(* IEC 61131-3 sources: daoli-st-library/DL_Motion (part 5) *)

(* ---- FB_DL_AgvPathTrackSeq.st ---- *)
// FB_DL_AgvPathTrackSeq v1.0.0
// 开源溯源：clean-room 自研（族 DL_Motion，ST 生态实测 0 命中，无外部代码引入）
(*
  功能: AGV 路径跟踪序列相位机：IDLE →(xStart∧xEnable) ALIGN →(双容差对齐) TRACK
        →(xObstacle) AVOID →(障碍解除∧保持 2 s) TRACK；TRACK →(xDockZone) DOCK
        →(对齐∧dist<0.05) IDLE 置 xDone。速度按 0.5 m/s² 斜坡逼近（增量 0.5·fCycleS，不阶跃），
        AVOID 与 FAULT 相强制零速零转。几何律全部委托外部 FC，本件不含三角函数。
  邻件: 对桩律 FC_DL_AgvChargeDockAlignCalc、限速 FC_DL_AgvSpeedLimitProfileCalc 为上游计算件。
  码表: 9311 入参非有限｜9312 组态非法(fSpeedLimit/fCycleS≤0)｜9313 相超时(ALIGN 5s/AVOID 保持/DOCK 15s)
        9314 相位落 ELSE 兜底｜9315 信息级序列完成（不置故障）。故障码锁存至 xReset 上升沿。
  边界: 无方法块/无属性块/无全局变量/无物理 IO 地址；三 TON 单相独占且无条件刷新。
*)
TYPE E_DL_AgvTrackState :
(
    IDLE  := 0,     // 空闲：等启动指令 [-] / Idle, waiting start
    ALIGN := 10,    // 对准：横向与角度对桩 [-] / Aligning to dock
    TRACK := 20,    // 跟踪：沿路径行驶 [-] / Tracking the path
    AVOID := 30,    // 避障：零速等待障碍解除 [-] / Avoiding obstacle
    DOCK  := 40,    // 入桩：末端贴近充电桩 [-] / Docking approach
    FAULT := 90     // 故障：锁存，仅复位沿可出 [-] / Fault latched
);
END_TYPE
FUNCTION_BLOCK FB_DL_AgvPathTrackSeq
VAR_INPUT
    xEnable     : BOOL := FALSE;        // 使能，FALSE 时全相冻结 [-] / Enable gate
    xStart      : BOOL := FALSE;        // 启动指令，上升沿有效 [-] / Start rising edge
    xReset      : BOOL := FALSE;        // 复位，上升沿清故障锁存 [-] / Reset rising edge
    xObstacle   : BOOL := FALSE;        // 障碍检测输入 [-] / Obstacle detected
    xDockZone   : BOOL := FALSE;        // 入桩区检测输入 [-] / Dock zone detected
    fOffsetY    : REAL := 0.0;          // 横向偏差 [m]，左正 / Lateral offset [m]
    fAngleErr   : REAL := 0.0;          // 角度偏差 [rad]，左正 / Angular error [rad]
    fDist       : REAL := 2.0;          // 到桩距离 [m] / Distance to dock [m]
    fSpeedLimit : REAL := 1.0;          // 允许限速 [m/s]，域 > 0 / Speed limit [m/s]
    fCycleS     : REAL := 0.01;         // 任务周期 [s]，域 > 0 / Task cycle time [s]
END_VAR
VAR_OUTPUT
    eState      : E_DL_AgvTrackState;   // 相位出口，段尾单点映射 [-] / Phase outlet
    xRun        : BOOL;                 // 运行中标志（非 IDLE 非 FAULT）[-] / Running flag
    fSpeedCmd   : REAL;                 // 前进速度指令 [m/s] / Speed command [m/s]
    fYawRateCmd : REAL;                 // 转向角速度指令 [rad/s] / Yaw rate command [rad/s]
    xDone       : BOOL;                 // 序列完成单拍脉冲 [-] / Done one-shot pulse
    xFault      : BOOL;                 // 故障锁存标志 [-] / Fault latch flag
    uErrorId    : UDINT;                // 事件码，0 = 无事件 / Event code
END_VAR
VAR
    tonAlign  : TON;                    // ALIGN 相超时 5 s，单相独占刷新 / Align timeout
    tonAvoid  : TON;                    // AVOID 障碍保持窗 2 s，单相独占刷新 / Avoid hold window
    tonDock   : TON;                    // DOCK 相超时 15 s，单相独占刷新 / Dock timeout
    rtStart   : R_TRIG;                 // 启动沿实例，无条件刷新 / Start edge instance
    rtReset   : R_TRIG;                 // 复位沿实例，无条件刷新 / Reset edge instance
    _eState   : E_DL_AgvTrackState := E_DL_AgvTrackState.IDLE;  // 内部相位，CASE 唯一写入 / Internal phase
    _fSpeed   : REAL := 0.0;            // 斜坡速度内部量 [m/s] / Ramp speed [m/s]
    _fSpTar   : REAL := 0.0;            // 本相速度目标 [m/s] / Phase speed target [m/s]
    _fYawTar  : REAL := 0.0;            // 本相转向目标 [rad/s] / Phase yaw target [rad/s]
    _fStep    : REAL := 0.0;            // 本周期斜坡增量 [m/s] / Per-cycle ramp step [m/s]
    _bAligned : BOOL := FALSE;          // 本拍对齐判据 [-] / Alignment judgement
    _bFault   : BOOL := FALSE;          // 故障锁存位（锁存量，仅复位沿清）/ Latched fault bit
    _uFault   : UDINT := 16#0000;       // 故障码锁存（锁存量，仅复位沿清）/ Latched fault code
    _uInfo    : UDINT := 16#0000;       // 信息码，每拍重算 / Transient info code
END_VAR
// 段 0：定时器与沿实例无条件周期刷新（禁置于 IF/CASE 内，R7）/ Unconditional refresh
rtStart(CLK := xStart);                                              // 启动沿每拍必调 / Start edge
rtReset(CLK := xReset);                                              // 复位沿每拍必调 / Reset edge
tonAlign(IN := (_eState = E_DL_AgvTrackState.ALIGN), PT := T#5S);    // 对准相超时 / Align timeout
tonAvoid(IN := (_eState = E_DL_AgvTrackState.AVOID), PT := T#2S);    // 避障保持窗 / Avoid window
tonDock(IN := (_eState = E_DL_AgvTrackState.DOCK), PT := T#15S);     // 入桩相超时 / Dock timeout
// 段 1：单拍量预清零（锁存量 _bFault/_uFault/_fSpeed 不入清单，R187）/ One-shot clear
_uInfo := 16#0000;                  // 信息码每拍重算 / Info code recomputed
xDone := FALSE;                     // 完成脉冲缺省清 / Done pulse clear
_fSpTar := 0.0;                     // 速度目标缺省零 / Speed target default zero
_fYawTar := 0.0;                    // 转向目标缺省零 / Yaw target default zero
_bAligned := FALSE;                 // 对齐判据缺省假 / Alignment default false
// 段 2：非有限闸与组态域闸（归因唯一，逐因独立码，R190）/ Gate stage
IF (fOffsetY <> fOffsetY) OR (fAngleErr <> fAngleErr) OR (fDist <> fDist)
   OR (fSpeedLimit <> fSpeedLimit) OR (fCycleS <> fCycleS)
   OR (ABS(fOffsetY) >= 3.0E38) OR (ABS(fAngleErr) >= 3.0E38) OR (ABS(fDist) >= 3.0E38)
   OR (ABS(fSpeedLimit) >= 3.0E38) OR (ABS(fCycleS) >= 3.0E38) THEN
    _uFault := 16#0002_9311;        // 故障级：入参非有限 / Fault: non-finite input
    _bFault := TRUE;                // 置故障锁存（R45 配对）/ Set fault latch
END_IF
IF (fSpeedLimit <= 1.0E-6) OR (fCycleS <= 1.0E-6) THEN
    _uFault := 16#0002_9312;        // 故障级：组态非法 / Fault: illegal configuration
    _bFault := TRUE;                // 置故障锁存（R45 配对）/ Set fault latch
END_IF
// 段 3：复位沿（FAULT 唯一解除路径）/ Reset edge, the only exit from fault
IF rtReset.Q THEN                   // rtReset.Q = 当拍量 / Reset edge is per-scan
    IF _eState = E_DL_AgvTrackState.FAULT THEN
        _eState := E_DL_AgvTrackState.IDLE;     // 故障相迁出回空闲 / Fault exits to idle
    END_IF
    _fSpeed := 0.0;                 // 斜坡量归零（锁存量解除）/ Ramp cleared on reset
    _bFault := FALSE;               // 清故障锁存位（仅此解除沿可清）/ Clear latched bit
    _uFault := 16#0000;             // 清故障锁存码（仅此解除沿可清）/ Clear latched code
END_IF
// 段 3b：对齐判据（ALIGN 与 DOCK 共用）/ Alignment judgement shared by two phases
IF (ABS(fOffsetY) <= 0.02) AND (ABS(fAngleErr) <= 0.03) THEN
    _bAligned := TRUE;              // 双容差内判对齐 / Within both tolerances
END_IF
// 段 4：相位机（本拍合法事件优先于超时，R275）/ Phase machine
CASE _eState OF
E_DL_AgvTrackState.IDLE:
    IF _bFault THEN
        _eState := E_DL_AgvTrackState.FAULT;        // 聚合故障进故障相 / Enter fault
    ELSIF rtStart.Q AND xEnable THEN
        _fSpeed := 0.0;                             // 起步斜坡复位 / Reset ramp on start
        _eState := E_DL_AgvTrackState.ALIGN;        // 进对准相 / Enter align
    END_IF
E_DL_AgvTrackState.ALIGN:
    IF _bFault THEN
        _eState := E_DL_AgvTrackState.FAULT;        // 故障优先 / Fault first
    ELSIF NOT xEnable THEN
        _eState := E_DL_AgvTrackState.IDLE;         // 使能撤销回空闲 / Enable dropped
    ELSIF _bAligned THEN
        _eState := E_DL_AgvTrackState.TRACK;        // 对齐到位进跟踪 / Aligned, track
    ELSIF tonAlign.Q THEN
        _uFault := 16#0002_9313;                    // 故障级：对准相超时 / Align timeout
        _bFault := TRUE;                            // 置故障锁存（R45 配对）/ Set latch
        _eState := E_DL_AgvTrackState.FAULT;        // 进故障相 / Enter fault
    ELSE
        IF fDist > 0.0 THEN
            _fSpTar := 0.3 * fDist;                 // 距离比例降速 / Distance speed
        ELSE
            _fSpTar := 0.0;                         // 距离为负/零：零速（R92 修，禁倒车指令）
        END_IF
        IF _fSpTar > 0.2 THEN
            _fSpTar := 0.2;                         // 对准相限速上限 / Align ceiling
        END_IF
        _fYawTar := 1.5 * fAngleErr;                // 角度比例转向 / Angular yaw
    END_IF
E_DL_AgvTrackState.TRACK:
    IF _bFault THEN
        _eState := E_DL_AgvTrackState.FAULT;        // 故障优先 / Fault first
    ELSIF NOT xEnable THEN
        _eState := E_DL_AgvTrackState.IDLE;         // 使能撤销回空闲 / Enable dropped
    ELSIF xObstacle THEN
        _eState := E_DL_AgvTrackState.AVOID;        // 障碍进避障 / Obstacle, avoid
    ELSIF xDockZone THEN
        _eState := E_DL_AgvTrackState.DOCK;         // 入桩区进入桩 / Dock zone, dock
    ELSE
        _fSpTar := fSpeedLimit;                     // 跟踪取限速 / Tracking uses limit
        _fYawTar := 1.0 * fAngleErr;                // 航向保持转向 / Heading hold yaw
    END_IF
E_DL_AgvTrackState.AVOID:
    IF NOT xEnable THEN
        _eState := E_DL_AgvTrackState.IDLE;         // 使能撤销回空闲 / Enable dropped
    ELSIF (NOT xObstacle) AND tonAvoid.Q THEN
        _eState := E_DL_AgvTrackState.TRACK;        // 障碍解除且保持到位回跟踪 / Cleared with hold
    ELSE
        _fSpeed := 0.0;                             // 避障零速（安全侧）/ Avoid zero speed
    END_IF
E_DL_AgvTrackState.DOCK:
    IF _bFault THEN
        _eState := E_DL_AgvTrackState.FAULT;        // 故障优先 / Fault first
    ELSIF NOT xEnable THEN
        _eState := E_DL_AgvTrackState.IDLE;         // 使能撤销回空闲 / Enable dropped
    ELSIF _bAligned AND (fDist < 0.05) THEN
        _fSpeed := 0.0;                             // 到位停稳 / Stop on position
        xDone := TRUE;                              // 完成脉冲单拍 / One-shot done
        _uInfo := 16#0002_9315;                     // 信息级：序列完成 / Info: done
        _eState := E_DL_AgvTrackState.IDLE;         // 回空闲 / Return to idle
    ELSIF tonDock.Q THEN
        _uFault := 16#0002_9313;                    // 故障级：入桩相超时 / Dock timeout
        _bFault := TRUE;                            // 置故障锁存（R45 配对）/ Set latch
        _eState := E_DL_AgvTrackState.FAULT;        // 进故障相 / Enter fault
    ELSE
        IF fDist > 0.0 THEN
            _fSpTar := 0.3 * fDist;                 // 末端贴近降速 / Final approach
        ELSE
            _fSpTar := 0.0;                         // 距离为负/零：零速（R92 修）
        END_IF
        IF _fSpTar > 0.1 THEN
            _fSpTar := 0.1;                         // 入桩相限速上限 / Dock ceiling
        END_IF
        _fYawTar := 1.5 * fAngleErr;                // 末段角度纠正 / Final angular fix
    END_IF
E_DL_AgvTrackState.FAULT:
    _fSpeed := 0.0;                                 // 故障相零速保持 / Fault zero speed
    IF rtReset.Q THEN
        _eState := E_DL_AgvTrackState.IDLE;         // 复位沿解除（段 3 已清锁存）/ Reset releases
    END_IF
ELSE
    _uFault := 16#0002_9314;                        // 故障级：非法相位兜底 / Illegal phase id
    _bFault := TRUE;                                // 置故障锁存（R45 配对）/ Set latch
    _fSpeed := 0.0;                                 // 非法相位零速 / Illegal phase zero speed
    _eState := E_DL_AgvTrackState.FAULT;            // 强制进故障相 / Force into fault
END_CASE
// 段 4b：转向目标限幅 ±0.4 rad/s / Yaw target clamping
IF _fYawTar > 0.4 THEN
    _fYawTar := 0.4;                                // 上饱和 / Upper saturation
ELSIF _fYawTar < -0.4 THEN
    _fYawTar := -0.4;                               // 下饱和 / Lower saturation
END_IF
// 段 4c：速度斜坡（禁阶跃；AVOID/FAULT 相不回填）/ Speed ramp, no step allowed
IF (_eState = E_DL_AgvTrackState.AVOID) OR (_eState = E_DL_AgvTrackState.FAULT) THEN
    _fSpeed := 0.0;                                 // 安全相斜坡归零 / Safety phases zero
ELSE
    _fStep := 0.5 * fCycleS;                        // 增量 = 0.5·fCycleS / Per-cycle step
    IF _fSpeed < _fSpTar THEN
        _fSpeed := _fSpeed + _fStep;                // 斜坡升速 / Ramp up
        IF _fSpeed > _fSpTar THEN
            _fSpeed := _fSpTar;                     // 不得越过目标 / No overshoot
        END_IF
    ELSIF _fSpeed > _fSpTar THEN
        _fSpeed := _fSpeed - _fStep;                // 斜坡降速 / Ramp down
        IF _fSpeed < _fSpTar THEN
            _fSpeed := _fSpTar;                     // 不得越过目标 / No overshoot
        END_IF
    END_IF
END_IF
// 段 5：出口单点映射（名实双出口，R191）/ Outlet mapping
eState := _eState;                                  // 相位出口单点映射 / Phase outlet
IF (_eState = E_DL_AgvTrackState.FAULT) OR _bFault THEN
    fSpeedCmd := 0.0;                               // 故障侧速度硬零 / Fault speed hard zero
    fYawRateCmd := 0.0;                             // 故障侧转向硬零 / Fault yaw hard zero
    xRun := FALSE;                                  // 故障侧非运行 / Not running
    xFault := TRUE;                                 // 故障锁存回放 / Replay latched flag
    uErrorId := _uFault;                            // 故障码锁存回放 / Replay latched code
ELSIF _eState = E_DL_AgvTrackState.IDLE THEN
    fSpeedCmd := 0.0;                               // 空闲相零速 / Idle zero speed
    fYawRateCmd := 0.0;                             // 空闲相零转 / Idle zero yaw
    xRun := FALSE;                                  // 空闲相非运行 / Not running
    xFault := FALSE;                                // 无故障 / No fault
    uErrorId := _uInfo;                             // 信息码重组 / Transient info code
ELSE
    fSpeedCmd := _fSpeed;                           // 运行相输出斜坡速度 / Ramp speed outlet
    fYawRateCmd := _fYawTar;                        // 运行相输出限幅转向 / Clamped yaw outlet
    xRun := TRUE;                                   // 运行中 / Running
    xFault := FALSE;                                // 无故障 / No fault
    uErrorId := _uInfo;                             // 信息码重组 / Transient info code
END_IF
IF (fSpeedCmd <> fSpeedCmd) OR (fYawRateCmd <> fYawRateCmd)
   OR (ABS(fSpeedCmd) >= 3.0E38) OR (ABS(fYawRateCmd) >= 3.0E38) OR (fSpeedCmd < 0.0) THEN
    fSpeedCmd := 0.0;                               // 出口复核失败回零速 / Outlet recheck zero
    fYawRateCmd := 0.0;                             // 出口复核失败回零转 / Outlet recheck zero
    xRun := FALSE;                                  // 复核失败撤运行 / Clear running
    xFault := TRUE;                                 // 复核失败置故障 / Raise fault
    uErrorId := 16#0002_9311;                       // 故障级：出口非有限 / Fault: non-finite outlet
END_IF
END_FUNCTION_BLOCK

(* ---- FB_DL_AxisAbortSafeSeq.st ---- *)
(*
  FB_DL_AxisAbortSafeSeq  —  运动中止安全序列（Abort→Stop→Disable 三段） / Axis abort safe sequence: stop, standstill wait, disable
  分类 Category : DL_Motion
  版本 Version  : 1.0.1
  来源 Source   : t1-6-plcopen — 运动序列族零检索深化（R233 成对纪律落地）
  溯源 Origin   : clean-room 实现，PLCopen 中止语义公开借鉴，未复制任何源码行
  功能 Function : 1) 三段顺控：eAbortStop（单发 iAxis.Stop，等轴受理反馈进
                  eStopping/eStandstill/eDisabled 稳态后迁出）→ eWaitStandstill
                  （等轴回 eStandstill）→ eDisable（单发 iAxis.Enable(bOn:=FALSE)，
                  等 bEnabled 落 FALSE）→ eDone；每段超时 TON 独立实例
                  （R233：配方推进与超时分件分实例）；
                  2) iAxis.bError → 故障级 03B1 锁存；段超时 → 03B2 锁存；
                  3) eFault 迁出边全当拍量（R240 落地），逐 BOOL 标注见段 5。
  返修记录 Rework  :
    2026-11-19  v1.0.1  R42 P0-4 轻度返修：v1.0.0 eAbortStop 相在单发 Stop 的
                        同拍即迁出 eWaitStandstill——该相驻留仅一个扫描拍，
                        tonStopTo 的 IN 只见单拍 TRUE，超时判据结构性不可达，
                        Stop 受理失败（轴拒收）将静默跳相（P0 派单缺陷④）。
                        修复要点：eAbortStop 相改为驻留等轴受理稳态
                        （eStopping/eStandstill/eDisabled 任一），受理确认后
                        才迁出；tonStopTo 跨相驻留恢复可计时性；对外接口
                        签名不变。
  边界 Boundary : ① 段迁出条件可满足性逐字自证：
                  eAbortStop → eWaitStandstill：Stop 受理后轴必进 eStopping（接口语义），
                  再至 eStandstill（受控停完成），迁出条件 eState 落已知稳态，可达；
                  eWaitStandstill → eDisable：轴停稳回 eStandstill 为接口规定稳态，可达；
                  eDisable → eDone：Enable(bOn:=FALSE) 后 bEnabled 落 FALSE 为接口规定
                  迁移（eStandstill → eDisabled），可达；
                  eFault 迁出：rtReset.Q AND NOT iAxis.bError AND bSrvOk（轴报警复位后 +
                  复位沿），可达；
                  ② 超时 TON 均单相独占（IN 为单相等式），跨相迁移拍 IN 必断（R228-A）；
                  ③ 组态闸：任一超时 <= 0 → 03B2 同级锁存（组态与超时归并为段超时码）；
                  ④ 无 GVL 依赖：纯引脚输入输出，无外部变量引用，无物理 IO 地址。
  依赖 Depends  : I_DL_MotionAxis（注入，不实例化）；Standard.library（TON / R_TRIG）
  码表 Error codes（Motion 段 0004，窗口 03B1~03B3 / 04B1~04B3）:
    16#0004_03B1 故障级：轴故障锁存（iAxis.bError），锁存至 bReset
    16#0004_03B2 故障级：段超时或组态非法（Abort/Wait/Disable 各相独立计时），锁存至 bReset
    16#0004_03B3 故障级：相位落 ELSE 兜底（非法相位 ID），锁存至 bReset
    16#0004_04B1 信息级：序列完成（eDone 相）
    16#0004_04B2 信息级：中止指令受理（Stop 单发拍）
    16#0004_04B3 信息级：使能切断确认（bEnabled 落 FALSE 拍）
  修订历史 Revision :
    2026-11-19  v1.0.0  R41 首版（批次 3 · 序号 2）
    2026-11-19  v1.0.1  R42 P0-4 轻度返修（见返修记录节）
*)

TYPE E_DL_AbsSeqState :
(
    eIdle            := 0,    // 空闲：等中止指令 / Idle, waiting abort command
    eAbortStop       := 10,   // 受停：单发 Stop，等轴受理 / Abort stop issued, waiting acceptance
    eWaitStandstill  := 20,   // 等停稳：等轴回 eStandstill / Waiting axis standstill
    eDisable         := 30,   // 切使能：单发 Enable(FALSE)，等 bEnabled 落 / Disable, waiting bEnabled off
    eDone            := 40,   // 完成：安全序列落定 / Done
    eFault           := 90    // 故障：轴故障/超时锁定 / Fault, latched
);
END_TYPE

FUNCTION_BLOCK FB_DL_AxisAbortSafeSeq
VAR_INPUT
    bAbortCmd    : BOOL := FALSE;     // 中止指令（上升沿启动序列）[-] / Abort command, starts on edge
    tStopTo      : TIME := T#2S;      // 受停相超时 [ms]，域 > 0 / Stop-phase timeout
    tStillTo     : TIME := T#10S;     // 等停稳相超时 [ms]，域 > 0 / Standstill-phase timeout
    tDisTo       : TIME := T#2S;      // 切使能相超时 [ms]，域 > 0 / Disable-phase timeout
    bReset       : BOOL := FALSE;     // 复位，上升沿清故障锁存（eFault 唯一迁出沿之一）/ Reset edge
END_VAR
VAR_IN_OUT
    iAxis        : I_DL_MotionAxis;   // 运动轴引用（注入，不实例化）/ Motion axis reference
END_VAR
VAR_OUTPUT
    eState       : E_DL_AbsSeqState;  // 状态出口，段尾单点映射 / State outlet
    bDone        : BOOL;              // 序列完成标志（eDone 相电平）/ Sequence done flag
    bCmdAccepted : BOOL;              // 中止指令受理单拍镜像 [-] / Command accepted mirror
    bError       : BOOL;              // 故障锁存标志 / Fault latch flag
    nErrId       : UDINT;             // 事件码，0 = 无事件 / Event code
END_VAR
VAR
    tonStopTo    : TON;               // 受停相超时（单相独占），无条件刷新 / Stop-phase timeout
    tonStillTo   : TON;               // 等停稳相超时（单相独占），无条件刷新 / Standstill timeout
    tonDisTo     : TON;               // 切使能相超时（单相独占），无条件刷新 / Disable-phase timeout
    rtAbort      : R_TRIG;            // 中止指令沿实例，无条件刷新 / Abort edge instance
    rtReset      : R_TRIG;            // 复位沿实例，无条件刷新 / Reset edge instance
    _eState      : E_DL_AbsSeqState := E_DL_AbsSeqState.eIdle;  // 内部相位（CASE 唯一写入目标）/ Internal phase
    _bCmdLatch   : BOOL;              // 本相命令已单发标志 / Phase command one-shot latch
    _bFault      : BOOL;              // 故障锁存位（锁存量）/ Latched fault bit
    _uFault      : UDINT;             // 故障码锁存（锁存量）/ Latched fault code
    _uInfo       : UDINT;             // 信息码，每拍重算 / Transient info code
END_VAR

(* —— 段 0：定时器与沿实例无条件周期刷新（禁置于 IF/CASE 内） —— *)
rtAbort(CLK := bAbortCmd);                                // 中止沿（每拍必调）
rtReset(CLK := bReset);                                   // 复位沿（每拍必调）
tonStopTo(IN := (_eState = E_DL_AbsSeqState.eAbortStop), PT := tStopTo);       // 受停超时（单相独占）
tonStillTo(IN := (_eState = E_DL_AbsSeqState.eWaitStandstill), PT := tStillTo); // 等停稳超时（单相独占）
tonDisTo(IN := (_eState = E_DL_AbsSeqState.eDisable), PT := tDisTo);           // 切使能超时（单相独占）

(* —— 段 1：单拍量预清零（锁存量 _bFault/_uFault 不入清单，禁同拍抹除） —— *)
_uInfo := 16#0000_0000;             // 信息码每拍重算
bCmdAccepted := FALSE;              // 受理镜像缺省 FALSE
nErrId := 16#0000_0000;             // 事件码缺省无事件

(* —— 段 2：轴故障与复位沿（判据当拍量） —— *)
IF iAxis.bError THEN                // iAxis.bError = 当拍量
    _uFault := 16#0004_03B1;        // 故障级：轴故障锁存
    _bFault := TRUE;
    iAxis.Stop();                   // 故障安全侧受控停
END_IF
IF (TIME_TO_DINT(tStopTo) <= 0) OR (TIME_TO_DINT(tStillTo) <= 0) OR (TIME_TO_DINT(tDisTo) <= 0) THEN
    _uFault := 16#0004_03B2;        // 故障级：组态非法（归并段超时码，头注释③）
    _bFault := TRUE;
END_IF
IF rtReset.Q AND (NOT iAxis.bError) THEN
(* 解除式逐 BOOL 标注（R240）：rtReset.Q = 当拍量；iAxis.bError = 当拍量；无锁存量自指。 *)
    IF _eState = E_DL_AbsSeqState.eFault THEN
        _eState := E_DL_AbsSeqState.eIdle;  // 故障相迁出：回空闲
    END_IF
    _bFault := FALSE;               // 清故障锁存位（锁存量，仅此当拍量解除沿可清）
    _uFault := 16#0000_0000;        // 清故障锁存码（锁存量，仅本当拍量解除沿可清）
END_IF

(* —— 段 3：相位机（只做迁移与单发命令；出口在段 5） —— *)
CASE _eState OF

E_DL_AbsSeqState.eIdle:
    IF rtAbort.Q AND (NOT _bFault) THEN
        _bCmdLatch := FALSE;                // 单发标志复位
        _eState := E_DL_AbsSeqState.eAbortStop;  // 进受停相
    END_IF

E_DL_AbsSeqState.eAbortStop:
    IF _bFault THEN
        _eState := E_DL_AbsSeqState.eFault; // 聚合故障直接进故障相
    ELSIF tonStopTo.Q THEN
        _uFault := 16#0004_03B2;            // 故障级：受停相超时（v1.0.1 相驻留承载，判据可达）
        _bFault := TRUE;
        _eState := E_DL_AbsSeqState.eFault;
    ELSE
        IF NOT _bCmdLatch THEN
            iAxis.Stop();                   // 单发受停命令（仅首拍）
            _bCmdLatch := TRUE;             // 单发标志
            _uInfo := 16#0004_04B2;         // 信息级：中止指令受理
            bCmdAccepted := TRUE;           // 受理镜像（单拍）
        END_IF
        IF (iAxis.eState = E_DL_AxisState.eStopping)         // 轴受理稳态 1：受控停中
           OR (iAxis.eState = E_DL_AxisState.eStandstill)    // 轴受理稳态 2：已停稳
           OR (iAxis.eState = E_DL_AxisState.eDisabled) THEN // 轴受理稳态 3：已失能
            _bCmdLatch := FALSE;                // 单发标志复位（下一相复用前）
            _eState := E_DL_AbsSeqState.eWaitStandstill;  // 受理确认：迁出（v1.0.1 驻留承载）
        END_IF
    END_IF

E_DL_AbsSeqState.eWaitStandstill:
    IF _bFault THEN
        _eState := E_DL_AbsSeqState.eFault; // 故障相
    ELSIF tonStillTo.Q THEN
        _uFault := 16#0004_03B2;            // 故障级：等停稳相超时
        _bFault := TRUE;
        _eState := E_DL_AbsSeqState.eFault;
    ELSE
        IF (iAxis.eState = E_DL_AxisState.eStandstill)
           OR (iAxis.eState = E_DL_AxisState.eDisabled) THEN
            _bCmdLatch := FALSE;            // 单发标志复位
            _eState := E_DL_AbsSeqState.eDisable;     // 停稳确认：进切使能相
        END_IF
    END_IF

E_DL_AbsSeqState.eDisable:
    IF _bFault THEN
        _eState := E_DL_AbsSeqState.eFault; // 故障相（使能请求已停发）
    ELSIF tonDisTo.Q THEN
        _uFault := 16#0004_03B2;            // 故障级：切使能相超时
        _bFault := TRUE;
        _eState := E_DL_AbsSeqState.eFault;
    ELSE
        IF NOT _bCmdLatch THEN
            iAxis.Enable(bOn := FALSE);     // 单发下使能命令
            _bCmdLatch := TRUE;             // 单发标志
        END_IF
        IF NOT iAxis.bEnabled THEN
            _uInfo := 16#0004_04B3;         // 信息级：使能切断确认
            _eState := E_DL_AbsSeqState.eDone;        // 进完成相
        END_IF
    END_IF

E_DL_AbsSeqState.eDone:
    bDone := TRUE;                      // 完成标志（eDone 相电平）
    _uInfo := 16#0004_04B1;             // 信息级：序列完成
    IF NOT bAbortCmd THEN
        bDone := FALSE;                 // 指令撤销：完成标志随相清除
        _eState := E_DL_AbsSeqState.eIdle;        // 回空闲
    END_IF

E_DL_AbsSeqState.eFault:
    ;                                   // 故障相：等复位沿（段 2 承载迁出）

ELSE
    _uFault := 16#0004_03B3;            // 故障级：非法相位 ID 兜底
    _bFault := TRUE;
    _eState := E_DL_AbsSeqState.eFault; // 强制回故障相

END_CASE

(* —— 段 4：出口单点映射（名实同源；锁存码回放，禁同拍抹除） —— *)
IF _bFault THEN
    nErrId := _uFault;              // 故障锁存码回放
    bDone := FALSE;                 // 故障相完成出口强制 FALSE（安全侧）
    bCmdAccepted := FALSE;          // 故障相受理镜像强制 FALSE（安全侧）
ELSE
    nErrId := _uInfo;               // 信息码
END_IF
bError := _bFault;                  // 故障标志与锁存位同源
eState := _eState;                  // 状态出口单点映射

END_FUNCTION_BLOCK

(* ---- FB_DL_AxisAccelFeedforward.st ---- *)
(*
  ==================================================================
  组件名 Component  : FB_DL_AxisAccelFeedforward
  分类   Category   : DL_Motion
  复杂度 Complexity  : cx3
  版本   Version    : 1.0.1
  功能   Purpose    : 轴加速度前馈注入。前馈叠加值 = Ka·aCmd + Kv·fVelAct，经一阶
                      低通平滑（滤波时间常数 fTauS）防抖后输出；bEnable 为假时
                      输出冻结保持并显式声明；参数（增益为负、周期非正、增益非
                      有限）一律回钳或判无效。
  来源   Source     : t1-6-plcopen
  溯源   Origin     : IEC 61131-3 标准语义的道莅防御性实现；加速度前馈偏置为公开
                      运动控制结构（规划加速度 × 折算增益），clean-room 自研实现，
                      未复制任何闭源代码行。
  平台   Platform   : 纯 IEC 61131-3（LREAL 运算，无私有库、无幂运算符、无定时器实例）
  作者   Author     : 道莅代码库 · PLC 编程专家（R56）
  ------------------------------------------------------------------
  边界 Boundary     :
                      一 本件只算前馈叠加值，不做限幅策略、不做轴使能仲裁（属主边界）；
                      二 bEnabled = FALSE 时输出冻结保持末值（R191 显式声明）；
                      三 输入非有限时输出安全侧归零并冻结滤波保持量（R127 常量安全侧）；
                      四 无全局变量、无外部变量声明、无物理地址寻址。
  输出契约 Output contract:
                      fFfOut 在有效拍为滤后前馈值；bEnabled 为本拍前馈有效指示；
                      eFault 为锁存回放（eCfgBad 组态非法 / eInputBad 本拍输入非有限）。
  修订记录 Revision  :
    2026-11-20  v1.0.0  R56 首版（批 2 · 序号 9）
    2026-11-21  v1.0.1  R57 返修：有效拍内补 eInputBad 信息级成因恢复撤销（对齐 TwoDofPid 段 10 范式）
  ==================================================================
*)

TYPE E_DL_AffFault :
(
    eNone     := 0, // 无成因 / no cause
    eCfgBad   := 1, // 组态非法：增益或周期越域（故障级，与 bError 配对）/ illegal config, gain or period out of domain
    eInputBad := 2  // 本拍指令加速度或实际速度非有限（信息级，输出归零）/ the command acceleration or the actual velocity is non finite this scan, the outlet is zeroed
);
END_TYPE

FUNCTION_BLOCK FB_DL_AxisAccelFeedforward
VAR_INPUT
    bEnable : BOOL := TRUE;   // 前馈使能，假时输出冻结保持 [-] / feedforward enable, false freezes the outlet
    bReset  : BOOL := FALSE;  // 复位上升沿清故障锁存与滤波保持 [-] / reset rising edge clears the fault latch and the filter holder
    aCmd    : LREAL := 0.0;   // 规划指令加速度 [单位每平方秒] / planned command acceleration [unit per square second]
    fVelAct : LREAL := 0.0;   // 实际速度 [单位每秒] / actual velocity [unit per second]
    fKa     : LREAL := 0.0;   // 加速度前馈增益（负值回钳零）[前馈每单位加速度] / acceleration feedforward gain, negatives clamp to zero [feedforward per unit acceleration]
    fKv     : LREAL := 0.0;   // 速度前馈增益（负值回钳零）[前馈每单位速度] / velocity feedforward gain, negatives clamp to zero [feedforward per unit velocity]
    fTauS   : LREAL := 0.02;  // 低通滤波时间常数 [秒]，0 = 直通 / low pass time constant [second], zero is a passthrough
    fDtS    : LREAL := 0.01;  // 调用周期 [秒]，域 大于零 / call period [second], domain above zero
END_VAR
VAR_OUTPUT
    fFfOut  : LREAL := 0.0;  // 前馈叠加值出口 [前馈单位] / the feedforward outlet [feedforward unit]
    bEnabled: BOOL := FALSE; // 本拍前馈有效指示 [-] / the feedforward valid indicator this scan
    bInvalid: BOOL := FALSE; // 本拍输出无效（归零或冻结）[-] / the outlet is void this scan
    eFault  : E_DL_AffFault := E_DL_AffFault.eNone; // 成因出口，锁存回放 [枚举] / cause outlet replayed from the latch [enum]
    bError  : BOOL := FALSE; // 故障锁存标志 [-] / fault latch flag
END_VAR
VAR
    rtReset : R_TRIG; // 复位沿检测，段 0 无条件刷新 / reset edge, refreshed unconditionally in segment zero
    _eFaulC : E_DL_AffFault := E_DL_AffFault.eNone; // 故障级成因，锁存至复位沿 / fault cause, latched until the reset edge
    _bFault : BOOL := FALSE; // 故障锁存位 [-] / fault latch bit
    _bInit  : BOOL := FALSE; // 首扫初始化完成标志（R310）/ first scan initialisation flag
    _bInOk  : BOOL := FALSE; // 本拍两输入均有限 [-] / both inputs are finite this scan
    _fKaUse : LREAL := 0.0;  // 钳定后的加速度增益 [前馈每单位加速度] / the clamped acceleration gain
    _fKvUse : LREAL := 0.0;  // 钳定后的速度增益 [前馈每单位速度] / the clamped velocity gain
    _fRaw   : LREAL := 0.0;  // 滤波前前馈值 [前馈单位] / the pre filter feedforward
    _fW     : LREAL := 0.0;  // 一阶低通权 [无量纲] / the first order weight
END_VAR

// 段 0｜沿检测无条件周期刷新（禁入分支）/ segment 0, unconditional refresh of the edge detector
rtReset(CLK := bReset); // 复位沿无条件刷新 / unconditional refresh of the reset edge

// 段 1｜首扫初始化（R310）/ segment 1, first scan initialisation
IF NOT _bInit THEN // 首扫一拍 / the very first scan
    _bInit := TRUE; // 置首扫完成标志 / raise the first scan flag
    _eFaulC := E_DL_AffFault.eNone; // 故障级成因清零 / clear the fault cause
    _bFault := FALSE; // 故障锁存清零 / clear the fault latch
END_IF

// 段 2｜复位沿作用域：清锁存 / 清滤波保持量（两项逐项声明）/ segment 2, reset edge scope declared item by item
IF rtReset.Q THEN // 复位沿 / the reset edge
    _bFault := FALSE; // 作用域一：清故障锁存 / scope one, clear the fault latch
    _eFaulC := E_DL_AffFault.eNone; // 作用域一：清故障级成因 / scope one, clear the fault cause
    fFfOut := 0.0; // 作用域二：出口归零 / scope two, the outlet is zeroed
END_IF

// 段 3｜组态域闸与参数回钳（R117 两级回退）/ segment 3, the configuration gate and the parameter clamps
_fKaUse := fKa; // 增益直通 / the gain passes through
_fKvUse := fKv; // 增益直通 / the gain passes through
IF (fKa <> fKa) OR ((fKa - fKa) <> (fKa - fKa)) OR (fKv <> fKv) OR ((fKv - fKv) <> (fKv - fKv)) OR (fDtS <= 0.0) OR (fDtS <> fDtS) OR (fTauS < 0.0) OR (fTauS <> fTauS) THEN // 增益或时间参数非有限 / a gain or a time parameter is non finite
    IF NOT _bFault THEN // 未锁存才迁移（防同拍抹除）/ migrate only while unlatched
        _bFault := TRUE; // 置故障锁存 / raise the fault latch
        _eFaulC := E_DL_AffFault.eCfgBad; // 故障级成因（R45 配对 bError）/ the fault cause paired with bError
    END_IF
END_IF
IF _fKaUse < 0.0 THEN // 加速度增益负值回钳零（一级回默认，R117）/ a negative gain clamps to the default zero
    _fKaUse := 0.0; // 钳到零 / clamp to zero
END_IF
IF _fKvUse < 0.0 THEN // 速度增益负值回钳零 / a negative gain clamps to zero
    _fKvUse := 0.0; // 钳到零 / clamp to zero
END_IF

// 段 4｜输入有限性闸 / segment 4, the input finiteness gate
_bInOk := (aCmd = aCmd) AND ((aCmd - aCmd) = (aCmd - aCmd)) AND (fVelAct = fVelAct) AND ((fVelAct - fVelAct) = (fVelAct - fVelAct)); // 两输入有限性 / finiteness of both inputs

// 段 5｜前馈计算与低通平滑 / segment 5, the feedforward computation and the low pass
IF (NOT _bInOk) OR _bFault OR (NOT bEnable) THEN // 非有限、故障或未使能 / non finite, faulted or disabled
    IF (NOT _bInOk) AND (NOT _bFault) THEN // 输入缺陷才记信息级成因（故障锁存优先回放，不覆盖故障码）/ only an input defect records the informational cause, never over a fault latch
        _eFaulC := E_DL_AffFault.eInputBad; // 信息级成因 / the informational cause
    END_IF
    bEnabled := FALSE; // 前馈无效指示 / the feedforward is not valid
    IF NOT bEnable THEN // 失能拍：冻结保持末值（R191 显式声明）/ the disabled scan holds the last value frozen
        bInvalid := FALSE; // 失能保持不算无效 / a disable is not an invalidity
    ELSE // 非有限或故障拍：输出安全侧归零（R127 常量）/ a non finite or faulted scan zeroes the outlet
        fFfOut := 0.0; // 输出归零 / the outlet is zeroed
        bInvalid := TRUE; // 置无效标志 / raise the invalid flag
    END_IF
ELSE // 有效拍 / the valid scan
    _fRaw := _fKaUse * aCmd + _fKvUse * fVelAct; // 前馈叠加原始值 / the raw feedforward composition
    IF fTauS > 0.0 THEN // 低通开启 / the low pass is on
        _fW := fDtS / (fDtS + fTauS); // 一阶低通权，除子为周期加时间常数已证大于零 / the first order weight with a proven divisor
        fFfOut := fFfOut + _fW * (_fRaw - fFfOut); // 低通推进（出口即保持量）/ advance the low pass, the outlet is the holder
    ELSE // 直通口径 / the passthrough
        fFfOut := _fRaw; // 原始值直出 / the raw value passes out
    END_IF
    bEnabled := TRUE; // 前馈有效指示 / the feedforward is valid
    bInvalid := FALSE; // 无效标志为假 / the invalid flag is false
    IF (_eFaulC = E_DL_AffFault.eInputBad) AND (NOT _bFault) THEN // 输入已恢复 / the input has recovered
        _eFaulC := E_DL_AffFault.eNone; // 信息级成因随恢复撤销（v1.0.1 返修，对齐 TwoDofPid 段 10 范式）/ the informational cause is revoked on recovery (v1.0.1 fix)
    END_IF
END_IF

// 段 6｜统一出口 / segment 6, the unified outlet
eFault := _eFaulC; // 成因出口锁存回放 / the cause outlet replayed from the latch
bError := _bFault; // 故障标志与锁存位同源 / the fault flag shares the latch source
END_FUNCTION_BLOCK

(* ---- FB_DL_AxisBacklashComp.st ---- *)
(*
  组件名 Component   : FB_DL_AxisBacklashComp
  子库 Sublibrary    : DL_Motion
  版本 Version       : 1.0.0
  兼容性 Platform    : CODESYS 3.5 / TwinCAT 3 / 汇川 InoProShop / Machine Expert（仅 Standard.library）
  功能 Function      : 轴反向间隙补偿：
                       1) 方向反转沿检测：速度指令符号越过零速死区即判换向（含迟滞），
                       反转沿承载补偿目标翻转；
                       2) 间隙学习值注入：补偿目标 = 方向符号 × 学习值 / 2（两侧各半程），
                       学习值越域（|学习值| > 上限）即冻结沿用上次域内值并告警锁存；
                       3) 补偿量注入按速率限幅爬升（fFeedRateMmS），不阶跃注入；
                       4) 非有限速度判输入非法，补偿冻结在当前值（安全侧）。
  边界 Boundary      : ① 本件只出补偿偏移量 fCompOffsetMm，由上层叠加到位置设定；
                       ② 学习值信任来源为学习工序（头注释声明信任边界：学习值由
                       间隙学习流程写入，本件只做域闸不回写）；
                       ③ 除法前置域闸：fGapMaxMm <= 0、fFeedRateMmS <= 0 判组态非法；
                       ④ 换向死区 fZeroVelEpsMmS 防零速附近符号抖动（迟滞口径）；
                       ⑤ 故障锁存解除唯一路径 = bReset 上升沿（输入引脚，恒可达）；
                       ⑥ 无全局变量引用、无外部变量声明、无物理地址寻址。
  依赖 Depends       : Standard.library（R_TRIG / F_TRIG）
  溯源 Origin        : 道莅自研 clean-room（参考 t1-6-plcopen 运动接口分类与参数域，
                       零代码行复制；与 FB_DL_BacklashCompensator 分工：那件为通用
                       丝杠间隙查表补偿，本件为轴域反转沿 + 学习值注入闭环件）
  码位 Code          : 16#04_0_A8
  码表 Error codes（Motion 格 04_0_A8，单轨：故障 0x02A8 / 信息 0x01A8）:
    16#0004_02A8 故障级：组态非法（间隙上限/爬升速率 <= 0）或学习值越域冻结或
                 速度非有限，锁存至 bReset 上升沿
    16#0004_01A8 信息级：换向补偿注入完成沿（爬升到位拍）
  修订历史 Revision  :
    2026-11-19  v1.0.0  R44 首版（批次 1 · 序号 5）
*)

TYPE E_DL_AbcState :
(
    eIdle  := 0,    // 空闲：未使能，补偿保持 / Idle, compensation held
    eRun   := 10,   // 运行：换向监视 + 补偿注入 / Running, reversal watch and injection
    eFault := 90    // 故障：组态/越域/非有限锁存 / Fault, latched
);
END_TYPE

FUNCTION_BLOCK FB_DL_AxisBacklashComp
VAR_INPUT
    bEnable       : BOOL;                  // 使能（电平），FALSE 时补偿保持 [-] / Enable
    bReset        : BOOL;                  // 上升沿清故障锁存 [-] / Reset edge
    fVelCmdMmS    : REAL;                  // 速度指令 [mm/s]，符号即方向 / Velocity command
    fLearnGapMm   : REAL;                  // 间隙学习值 [mm]，学习工序写入 / Learned backlash value
    fGapMaxMm     : REAL := 0.5;           // 学习值域上限 [mm] / Learned value ceiling
    fZeroVelEpsMmS: REAL := 1.0;           // 换向零速死区 [mm/s] / Reversal zero-speed deadband
    fFeedRateMmS  : REAL := 10.0;          // 补偿注入爬升速率 [mm/s] / Injection slew rate
    tCycle        : TIME := T#10MS;        // 扫描周期 [毫秒] / Scan cycle time
END_VAR
VAR_OUTPUT
    fCompOffsetMm : REAL;                  // 补偿偏移量输出 [mm]，叠加到位置设定 / Compensation offset
    fGapUseMm     : REAL;                  // 生效学习值（域内钳用）[mm] / Effective learned gap
    bReversing    : BOOL;                  // 换向注入进行中电平 [-] / Reversal injection active
    bGapFrozen    : BOOL;                  // 学习值冻结标志 [-] / Learned value frozen flag
    eState        : E_DL_AbcState;         // 状态出口，段尾单点映射 / State outlet
    bError        : BOOL;                  // 故障锁存标志 [-] / Fault latch flag
    uErrId        : UDINT;                 // 事件码，0 = 无事件 / Event code
END_VAR
VAR
    rtReset   : R_TRIG;                    // 复位沿实例，段 0 无条件刷新 / Reset edge
    rtRevFwd  : R_TRIG;                    // 正向进入沿实例，段 0 无条件刷新 / Forward entry edge
    ftRevBwd  : F_TRIG;                    // 正向退出（反向进入）沿实例，段 0 无条件刷新 / Reverse entry edge
    _eState   : E_DL_AbcState := E_DL_AbcState.eIdle;   // 内部相位（CASE 唯一写入目标）/ Internal phase
    _bDirPos  : BOOL;                      // 方向电平（迟滞后）[-] / Direction level with hysteresis
    _fTarget  : REAL;                      // 补偿目标偏移 [mm] / Compensation target
    _fStep    : REAL;                      // 本拍注入步长 [mm] / Injection step per scan
    _bDirSeen : BOOL;                      // 首个有效方向已建立标志 [-] / First direction established
    _bFault   : BOOL;                      // 故障锁存位（锁存量） / Latched fault bit
    _uFault   : UDINT;                     // 故障码锁存（锁存量） / Latched fault code
    _bCfgBad  : BOOL;                      // 组态非法当拍量 [-] / Config illegal flag
    _bNonFin  : BOOL;                      // 输入非有限当拍量 [-] / Non-finite input flag
    _bInjDone : BOOL;                      // 注入到位当拍量 [-] / Injection settled flag
    _bReversingCalc : BOOL;                // 换向注入进行中内部量 [-] / Reversal injection internal
END_VAR
VAR CONSTANT
    DL_TWO     : REAL := 2.0;              // 半程系数（两侧各分半）[无量纲] / Half factor
    DL_STEP_EPS: REAL := 1.0E-9;           // 注入到位判据 [mm] / Injection settled tolerance
    DL_ABS_MAX : REAL := 1.0E30;           // 有限值判定上界 [mm] / Finite value bound
    DL_ZERO    : REAL := 0.0;              // 零常量 [mm] / Zero constant
    DL_MS_PER_S: REAL := 1000.0;           // 毫秒 → 秒换算系数 [毫秒/秒] / Milliseconds per second
END_VAR

(* —— 段 0｜沿实例每拍无条件刷新（禁置于 IF/CASE 内） —— *)
rtReset (CLK := bReset);
rtRevFwd(CLK := _bDirPos);
ftRevBwd(CLK := _bDirPos);

(* —— 段 1｜瞬时量预清零与周期换算（锁存量 _bFault/_uFault/fCompOffsetMm 不入清单） —— *)
uErrId   := 16#0000_0000;
_bCfgBad := FALSE;
_bNonFin := FALSE;
_bInjDone := FALSE;
_bReversingCalc := FALSE;

(* —— 段 2｜复位沿：故障一次性清干净，相位回空闲 —— *)
IF rtReset.Q THEN
    _bFault := FALSE;
    _uFault := 16#0000_0000;
    _eState := E_DL_AbcState.eIdle;
END_IF

(* —— 段 3｜组态闸与非有限判据（覆盖全部参与换算引脚） —— *)
IF (fGapMaxMm <= DL_ZERO) OR (fFeedRateMmS <= DL_ZERO) OR (fZeroVelEpsMmS <= DL_ZERO)
   OR (tCycle = T#0S) THEN
    _bCfgBad := TRUE;
END_IF
IF (fVelCmdMmS <> fVelCmdMmS) OR ((fVelCmdMmS - fVelCmdMmS) <> DL_ZERO)
   OR (fLearnGapMm <> fLearnGapMm) OR ((fLearnGapMm - fLearnGapMm) <> DL_ZERO) THEN
    _bNonFin := TRUE;
END_IF

(* —— 段 4｜主状态机：三态全覆盖 + ELSE 兜底 —— *)
CASE _eState OF

E_DL_AbcState.eIdle:
    IF bEnable AND (NOT _bCfgBad) AND (NOT _bNonFin) THEN
        bGapFrozen := FALSE;
        fGapUseMm  := ABS(fLearnGapMm);  // 首次进入按当下学习值启用
        _bDirSeen  := FALSE;
        _eState    := E_DL_AbcState.eRun;
    ELSIF bEnable AND (_bCfgBad OR _bNonFin) THEN
        _bFault := TRUE;                 // 故障级配对置位（R45）
        _uFault := 16#0004_02A8;
        bError  := TRUE;
        _eState := E_DL_AbcState.eFault;
    END_IF

E_DL_AbcState.eRun:
    IF NOT bEnable THEN
        _eState := E_DL_AbcState.eIdle;  // 使能撤销回空闲，补偿量保持
    ELSE
        (* 学习值域闸：越域即冻结沿用域内值，锁存告警 *)
        IF ABS(fLearnGapMm) > fGapMaxMm THEN
            bGapFrozen := TRUE;          // 冻结标志（锁存，复位沿解除）
            _bFault := TRUE;
            _uFault := 16#0004_02A8;
            bError  := TRUE;
            _eState := E_DL_AbcState.eFault;
        ELSE
            fGapUseMm := ABS(fLearnGapMm);   // 域内学习值照常更新
            bGapFrozen := FALSE;
        END_IF
        IF NOT _bFault THEN
            (* 换向判定：零速死区迟滞，防零速附近符号抖动 *)
            IF (NOT _bDirPos) AND (fVelCmdMmS > fZeroVelEpsMmS) THEN
                _bDirPos := TRUE;
                _bDirSeen := TRUE;
            ELSIF _bDirPos AND (fVelCmdMmS < -fZeroVelEpsMmS) THEN
                _bDirPos := FALSE;
                _bDirSeen := TRUE;
            END_IF
            IF _bDirSeen THEN
                IF _bDirPos THEN
                    _fTarget := fGapUseMm / DL_TWO;      // 正向：+半程
                ELSE
                    _fTarget := -fGapUseMm / DL_TWO;     // 反向：-半程
                END_IF
            ELSE
                _fTarget := DL_ZERO;     // 首方向未建立：目标归零
            END_IF
            (* 速率限幅注入：步长 = 速率 × 周期，不阶跃 *)
            _fStep := fFeedRateMmS * TIME_TO_REAL(tCycle) / DL_MS_PER_S;
            IF fCompOffsetMm < _fTarget THEN
                fCompOffsetMm := MIN(fCompOffsetMm + _fStep, _fTarget);
                _bReversingCalc := TRUE;
            ELSIF fCompOffsetMm > _fTarget THEN
                fCompOffsetMm := MAX(fCompOffsetMm - _fStep, _fTarget);
                _bReversingCalc := TRUE;
            ELSE
                _bInjDone := TRUE;       // 注入到位
            END_IF
            IF _bInjDone AND (rtRevFwd.Q OR ftRevBwd.Q) THEN
                uErrId := 16#0004_01A8;  // 信息级：换向注入完成沿
            END_IF
        END_IF
    END_IF

E_DL_AbcState.eFault:
    bError := TRUE;                      // 故障相驻留：补偿量冻结保持，只认复位沿（段 2 迁出）
    ;                                    // （冻结语义：fCompOffsetMm 保持最后值，安全侧不归零）

ELSE
    _bFault := TRUE;                     // 兜底：非法相位锁存
    _uFault := 16#0004_02A8;
    bError  := TRUE;
    _eState := E_DL_AbcState.eFault;
END_CASE

(* —— 段 5｜状态出口单点映射（名实同源） —— *)
bReversing := _bReversingCalc;           // 换向注入电平同源赋值（R191）
eState := _eState;
END_FUNCTION_BLOCK

(* ---- FB_DL_AxisBacklashStepComp.st ---- *)
(*
  Name        : FB_DL_AxisBacklashStepComp
  Category    : DL_Motion
  Version     : 1.0.1
  Purpose     : 轴反向间隙阶跃补偿：跟踪位置命令方向，方向切换拍一次性注入补偿行程（新方向补偿量累加到偏置），输出补偿后位置；/ Axis backlash step compensation: tracks command direction and injects the compensation travel as a one-shot step on each reversal by accumulating the offset into the commanded position
  溯源        : 借 t1-6-plcopen-motion 的分类/参数域组织，clean-room 实现
  Changelog   : v1.0.1 R54 非有限拍 fPosOut 直算 NaN 修复：出口计算移入有限分支，非有限拍保持上拍 fPosOut/fOffset 并置 bInvalid 当拍指示
  撞名说明    : 本件原名 FB_DL_AxisBacklashComp 与既有 R44 件（DL_Motion，换向沿 + 学习值注入 +
                速率爬升口径）撞名，为免 POU/枚举/常量三重重复定义，改名 FB_DL_AxisBacklashStepComp，
                枚举前缀 E_DL_AbsStep*、常量前缀 DL_ABS_ 全部隔离；分工：R44 件为速度指令口径的
                学习值爬升注入，本件为位置命令口径的方向切换拍阶跃注入。
  Boundary    : ① 组态闸：补偿量 < 0 → 锁存故障（0 = 关闭补偿，合法）；
                ② 方向判定：命令增量绝对值 > 判向阈才更新方向（死区防噪声反复触发注入）；
                ③ 注入只在方向切换当拍发生一次（沿语义），同向运行不重复注入；
                ④ 偏置饱和上限防 REAL 有效位耗尽（R28）；bCompPuls 单拍脉冲经内部 _b* 统一出口映射（R187）；
                ⑤ 非有限命令该拍不判向不注入（偏置与输出保持上拍值，防污染）；
                ⑥ 本件为映射层补偿，不替代驱动器内置补偿、不做安全限位（属主边界）。
*)
TYPE E_DL_AbsStepState :
(
    eIdle  := 0,                             (* 未使能 / Disabled *)
    eRun   := 10,                            (* 补偿跟踪运行 / Compensating *)
    eFault := 90                             (* 故障锁存相 / Fault latched *)
);
END_TYPE

TYPE E_DL_AbsStepCause :
(
    eNone       := 0,                        (* 无故障成因 / No cause *)
    eCfgIllegal := 1,                        (* 组态非法：补偿量为负 / Illegal config *)
    ePhaseBad   := 2                         (* 非法相位兜底 / Illegal phase fallback *)
);
END_TYPE

FUNCTION_BLOCK FB_DL_AxisBacklashStepComp
VAR_INPUT
    fPosCmd  : REAL := 0.0;                  (* 位置命令输入 [mm] / Command position input *)
    fBacklash: REAL := 0.02;                 (* 反向间隙补偿量，域 >= 0（0 = 关闭补偿）[mm] / Backlash compensation, >= 0 *)
    bEnable  : BOOL := TRUE;                 (* 补偿使能 [-] / Enable *)
    bReset   : BOOL := FALSE;                (* 复位命令，上升沿清偏置与故障 [-] / Reset command *)
END_VAR
VAR_OUTPUT
    fPosOut  : REAL;                         (* 补偿后位置输出 = 命令 + 偏置 [mm] / Compensated position output *)
    fOffset  : REAL;                         (* 当前累计偏置（镜像）[mm] / Current accumulated offset mirror *)
    bCompPuls: BOOL;                         (* 本拍发生方向切换注入（单拍脉冲）[-] / Injection this scan pulse *)
    nCompCnt : UDINT;                        (* 累计注入次数（诊断，饱和）[次] / Injection count, saturated *)
    bInvalid : BOOL;                         (* 命令非有限当拍指示（出口保持上拍值，v1.0.1）[-] / Non-finite command indicator *)
    eState   : E_DL_AbsStepState;            (* 状态出口 / State outlet *)
    eCause   : E_DL_AbsStepCause;            (* 故障成因出口（R190 归因唯一） / Fault cause outlet *)
    bError   : BOOL;                         (* 故障锁存标志 [-] / Fault latch flag *)
END_VAR
VAR
    _eState  : E_DL_AbsStepState := E_DL_AbsStepState.eIdle;    (* 内部相位（CASE 唯一写入目标） / Internal phase *)
    _eCause  : E_DL_AbsStepCause := E_DL_AbsStepCause.eNone;    (* 故障成因锁存量 / Latched cause *)
    rtReset  : R_TRIG;                       (* 复位沿实例，段 0 无条件调用 / Reset edge instance *)
    _bFault  : BOOL;                         (* 故障锁存位 / Latched fault bit *)
    _bCfgBad : BOOL;                         (* 组态非法当拍量 / Illegal config this scan *)
    _bFin    : BOOL;                         (* 位置命令有限性当拍量 / Command finiteness *)
    _bDirC   : BOOL;                         (* 方向切换注入内部单拍量（出口统一映射，R187） / Injection internal pulse *)
    _bBadI   : BOOL;                         (* 非有限命令当拍指示内部量（统一出口映射，R187，v1.0.1） / Invalid internal pulse *)
    _nDir    : INT := 0;                     (* 当前方向（+1 正 / -1 负 / 0 未定）[-] / Current direction *)
    _fPrev   : REAL;                         (* 上拍命令位置快照 [mm] / Previous command snapshot *)
    _fOffI   : REAL;                         (* 累计偏置内部量（fPosOut 的加数）[mm] / Accumulated offset internal *)
    _fDeltaI : REAL;                         (* 命令增量中间量 [mm] / Command delta intermediate *)
END_VAR
VAR CONSTANT
    DL_ABS_EPS    : REAL  := 1.0E-6;         (* 判零容差 [-] / Epsilon *)
    DL_ABS_DIRTH  : REAL  := 0.001;          (* 判向阈：增量绝对值超过此值才更新方向 [mm] / Direction threshold *)
    DL_ABS_OFFMAX : REAL  := 1.0E6;          (* 偏置饱和上限（防 REAL 有效位耗尽，R28）[mm] / Offset saturation cap *)
    DL_ABS_CNTMAX : UDINT := 4294967295;     (* 注入计数饱和上限（R28）[-] / Injection count cap *)
    DL_ABS_PLUS   : INT   := 1;              (* 正方向枚举值 [-] / Positive direction *)
    DL_ABS_MINUS  : INT   := -1;             (* 负方向枚举值 [-] / Negative direction *)
    DL_ABS_UNDEF  : INT   := 0;              (* 未定向值 [-] / Undefined direction *)
END_VAR

(* —— 段 0：当拍判据派生 + 实例无条件刷新（R228A） —— *)
_bCfgBad := (fBacklash < 0.0);                                                 (* 补偿量非负闸（0 = 关闭补偿合法） / Backlash non-negative gate *)
rtReset(CLK := bReset);                                                        (* 复位沿每拍必调 / Reset edge every scan *)
_bFin := (fPosCmd = fPosCmd) AND ((fPosCmd - fPosCmd) = (fPosCmd - fPosCmd));  (* 命令 NaN 自反 + Inf 差判闸 / Command NaN and Inf gate *)
_fDeltaI := 0.0;                                                               (* 增量中间量预置（非有限拍为 0 不判向） / Delta preset zero *)
IF _bFin AND (_eState = E_DL_AbsStepState.eRun) THEN
    _fDeltaI := fPosCmd - _fPrev;                                              (* 命令增量（运行相才派生）[mm] / Command delta in run phase *)
END_IF

(* —— 段 1：单拍量预清零（R107） —— *)
_bDirC := FALSE;                                                               (* 注入脉冲内部量预清 / Injection preset *)
_bBadI := FALSE;                                                               (* 非有限指示内部量预清（v1.0.1） / Invalid preset *)
bCompPuls := FALSE;                                                            (* 注入脉冲出口预清 / Injection outlet preset *)
bInvalid := FALSE;                                                             (* 非有限指示出口预清（v1.0.1） / Invalid outlet preset *)

(* —— 段 2：复位沿处理（作用域：清故障 + 清偏置与方向 + 迁 eIdle，R283 逐项声明） —— *)
IF rtReset.Q THEN
    _bFault := FALSE;                                                          (* 清故障锁存 / Clear fault *)
    _eCause := E_DL_AbsStepCause.eNone;                                        (* 清成因 / Clear cause *)
    _fOffI := 0.0;                                                             (* 清偏置内部量 / Clear offset internal *)
    fOffset := 0.0;                                                            (* 清偏置镜像出口 / Clear offset mirror *)
    fPosOut := 0.0;                                                            (* 清位置输出出口 / Clear position outlet *)
    bInvalid := FALSE;                                                         (* 清非有限指示出口（v1.0.1） / Clear invalid outlet *)
    nCompCnt := 0;                                                             (* 清注入计数出口 / Clear injection count *)
    _nDir := DL_ABS_UNDEF;                                                     (* 方向回未定 / Direction undefined *)
    _fPrev := 0.0;                                                             (* 清上拍快照 / Clear previous snapshot *)
    _eState := E_DL_AbsStepState.eIdle;                                        (* 迁未使能相 / Back to idle *)
END_IF

(* —— 段 3：组态故障锁存（锁存至复位沿，R189） —— *)
IF _bCfgBad AND NOT _bFault THEN
    _bFault := TRUE;                                                           (* 锁存故障位 / Latch fault *)
    _eCause := E_DL_AbsStepCause.eCfgIllegal;                                  (* 成因：组态非法 / Cause: illegal config *)
    _eState := E_DL_AbsStepState.eFault;                                       (* 同步迁故障相 / Migrate to fault *)
END_IF

(* —— 段 4：CASE 主状态机（ELSE 兜底迁 eFault，红线 6） —— *)
CASE _eState OF
    E_DL_AbsStepState.eIdle:                                                   (* 未使能：出口确定值 / Disabled *)
        fPosOut := 0.0;                                                        (* 失能清位置输出出口 / Clear position outlet *)
        fOffset := 0.0;                                                        (* 失能清偏置镜像出口 / Clear offset mirror *)
        bCompPuls := FALSE;                                                    (* 失能清注入脉冲出口 / Clear injection outlet *)
        _fOffI := 0.0;                                                         (* 失能清偏置内部量（防隐性回夹） / Clear offset internal *)
        _nDir := DL_ABS_UNDEF;                                                 (* 失能方向回未定（重使能重新定向） / Direction undefined *)
        IF bEnable AND NOT _bFault THEN
            _fPrev := fPosCmd;                                                 (* 迁入拍取命令首快照（首次增量不误判向） / Command snapshot at entry *)
            _eState := E_DL_AbsStepState.eRun;                                 (* 使能进入补偿 / Enter compensating *)
        END_IF
    E_DL_AbsStepState.eRun:                                                    (* 补偿相：判向 + 切换拍注入 / Compensating *)
        IF NOT bEnable THEN
            _eState := E_DL_AbsStepState.eIdle;                                (* 失能回未使能 / Back to idle *)
        ELSE
            IF _bFin THEN
                IF ABS(_fDeltaI) > DL_ABS_DIRTH THEN                           (* 增量超判向阈才更新方向（死区防噪声，边界②） / Direction update above threshold *)
                    IF _fDeltaI > 0.0 THEN
                        IF _nDir = DL_ABS_MINUS THEN                           (* 负 → 正方向切换：注入正补偿 / Reversal to positive *)
                            _bDirC := TRUE;                                    (* 注入脉冲内部置位（R187） / Injection internal *)
                            IF _fOffI < DL_ABS_OFFMAX THEN
                                _fOffI := _fOffI + fBacklash;                  (* 偏置累加补偿量（饱和防有效位耗尽） / Offset accumulate, capped *)
                            END_IF
                            IF nCompCnt < DL_ABS_CNTMAX THEN
                                nCompCnt := nCompCnt + 1;                      (* 注入计数净额 +1（饱和） / Net +1, saturated *)
                            END_IF
                        END_IF
                        _nDir := DL_ABS_PLUS;                                  (* 更新为正方向 / Set positive *)
                    ELSIF _fDeltaI < 0.0 THEN
                        IF _nDir = DL_ABS_PLUS THEN                            (* 正 → 负方向切换：注入负补偿 / Reversal to negative *)
                            _bDirC := TRUE;                                    (* 注入脉冲内部置位（R187） / Injection internal *)
                            IF _fOffI > -DL_ABS_OFFMAX THEN
                                _fOffI := _fOffI - fBacklash;                  (* 偏置累减补偿量（对称饱和） / Offset accumulate negative, capped *)
                            END_IF
                            IF nCompCnt < DL_ABS_CNTMAX THEN
                                nCompCnt := nCompCnt + 1;                      (* 注入计数净额 +1（饱和） / Net +1, saturated *)
                            END_IF
                        END_IF
                        _nDir := DL_ABS_MINUS;                                 (* 更新为负方向 / Set negative *)
                    END_IF
                END_IF
                _fPrev := fPosCmd;                                             (* 每拍刷新命令快照（有限拍才刷） / Refresh snapshot on finite scan *)
                fOffset := _fOffI;                                             (* 偏置镜像出口（有限拍才派生，v1.0.1 移入） / Offset mirror outlet *)
                fPosOut := fPosCmd + _fOffI;                                   (* 补偿后位置输出（有限拍才派生，v1.0.1 修复 NaN 穿透） / Compensated output *)
            ELSE
                _bBadI := TRUE;                                                (* 非有限拍：置失效指示内部量（R187，v1.0.1） / Invalid internal *)
            END_IF                                                             (* 非有限拍：不判向不注入，fPosOut/fOffset 保持上拍值（边界⑤） *)
        END_IF
    E_DL_AbsStepState.eFault:                                                  (* 故障相：冻结保持末值，仅复位沿出 / Fault *)
        ;                                                                      (* 锁存回放（R28） / Replay from latch *)
    ELSE                                                                       (* 非法相位兜底迁安全态 / Illegal phase fallback *)
        _eState := E_DL_AbsStepState.eFault;                                   (* 迁故障相 / To fault *)
        _bFault := TRUE;                                                       (* 同步锁存 / Latch *)
        _eCause := E_DL_AbsStepCause.ePhaseBad;                                (* 成因：非法相位 / Cause: illegal phase *)
END_CASE

(* —— 段 5：出口映射（内部 _b* → 输出单拍，R187；名实双出口，R191） —— *)
bCompPuls := _bDirC;                                                           (* 注入脉冲单拍出口 / Injection single-scan outlet *)
bInvalid := _bBadI;                                                            (* 非有限指示单拍出口（v1.0.1） / Invalid single-scan outlet *)
bError := _bFault;                                                             (* 故障标志镜像 / Fault flag mirror *)
eState := _eState;                                                             (* 状态出口 / State outlet *)
eCause := _eCause;                                                             (* 成因出口 / Cause outlet *)
END_FUNCTION_BLOCK

(* ---- FB_DL_AxisBrakeDistPredict.st ---- *)
(*
  FB_DL_AxisBrakeDistPredict  —  轴制动距离预判（速度/减速度→停车距离 + 硬限位留量） / Axis braking-distance prediction from velocity and deceleration with hard-limit allowance
  分类 Category : DL_Motion
  版本 Version  : 1.0.0
  来源 Source   : t1-6-plcopen — PLCopen Motion 接口映射层族深化
  溯源 Origin   : 道莅 clean-room 实现；匀减速停车距离 d = v×t_react + v²/(2a) 为公开运动学公式，
                 本件仅做 PLCopen MC 接口的判据映射层，不内联任何轨迹规划内核（复用 DL_Algo 既有件）
  功能 Function : 1) 反应距离 _fReactMm = fActVelMmS × 反应时间(s)；
                  2) 制动距离 _fBrakeMm = v² / (2 × fDecelMmS2)（除零前置判，减速度 <= 1.0E-6 判组态非法）；
                  3) 停车总距离 _fStopMm = 反应距离 + 制动距离 + fSafetyMarginMm；
                  4) 可用距离按运动方向取（正向 = 限位 - 当前；反向 = 当前 - 限位），负值钳制 0；
                  5) 判据：可用距离 > 停车总距离 → bStopOk；否则进 eBrake 相请求减速停车；
                  6) 本件只有故障码、无信息码（派单硬约束）。
  接口 Interface: 输入速度/减速度/位置/限位/余量/反应时间/方向；输出停车距离与判据
  边界 Boundary : ① 组态闸：fDecelMmS2 <= 1.0E-6、tReaction <= T#0S、fSafetyMarginMm < 0.0
                  → 04A6 锁存；② 速度/位置/限位非有限（NaN 自反 + Inf 差值自减）→ 04A6 锁存，
                  判据取安全侧（bStopOk = FALSE，请求停车）；
                  ③ 除零防护在计算前以减速度正域判据完成（不进入除法）；
                  ④ 一个 R_TRIG，段 0 无条件调用；⑤ 故障相迁出唯一路径 = bReset 上升沿；
                  ⑥ 零全局耦合：无 GVL / VAR_EXTERNAL / %I %Q %M 直接地址。
  依赖 Depends  : Standard.library（R_TRIG）
  码表 Error codes（Motion 段 0004，故障窗口 04A6；本件无信息码）:
    16#0004_04A6 故障级：制动距离预判故障总码（组态非法 / 输入非有限），
                 锁存至 bReset 上升沿；归因见 eCause，不新增码位（派单硬约束单码）
  修订历史 Revision :
    2026-11-19  v1.0.0  R43 首版（批次 4 · 序号 18）
*)

TYPE E_DL_AbpState :
(
    eIdle  := 0,      // 未使能待预判 / Idle, waiting prediction
    eRun   := 10,     // 预判运行中（距离充足） / Predicting, distance sufficient
    eBrake := 20,     // 距离不足：请求减速停车 / Insufficient distance, stop requested
    eFault := 90      // 故障锁存相（请求停车） / Fault latched, stop requested
);
END_TYPE

TYPE E_DL_AbpCause :
(
    eNone       := 0, // 无故障成因 / No cause
    eCfgIllegal := 1, // 组态非法 / Illegal configuration
    eNonFinite  := 2  // 输入非有限 / Non-finite input
);
END_TYPE

FUNCTION_BLOCK FB_DL_AxisBrakeDistPredict
VAR_INPUT
    fActVelMmS     : REAL := 0.0;      // 轴实际速度 [mm/s]，域 >= 0 / Actual axis velocity
    fDecelMmS2     : REAL := 1000.0;   // 规划减速度 [mm/s²]，域 > 0 / Planned deceleration
    fPosMm         : REAL := 0.0;      // 当前轴位置 [mm] / Current axis position
    fLimitPosMm    : REAL := 0.0;      // 硬限位位置 [mm] / Hard limit position
    fSafetyMarginMm: REAL := 10.0;     // 安全留量 [mm]，域 >= 0 / Safety margin
    tReaction      : TIME := T#50MS;   // 反应时间 [ms]，域 > 0 / Reaction time
    bDirPositive   : BOOL := TRUE;     // 运动方向：TRUE = 正向 [-] / Direction, TRUE = positive
    bEnable        : BOOL := FALSE;    // 预判使能（电平）[-] / Prediction enable
    bReset         : BOOL := FALSE;    // 复位命令，上升沿清故障 [-] / Reset edge
END_VAR
VAR_OUTPUT
    eState         : E_DL_AbpState;    // 状态出口，段 6 单点映射 / State outlet
    eCause         : E_DL_AbpCause;    // 故障成因出口（R190） / Fault cause outlet
    fStopDistMm    : REAL;             // 停车总距离 [mm] / Total stopping distance
    fAvailMm       : REAL;             // 到限位可用距离 [mm] / Available distance to limit
    bStopOk        : BOOL;             // 距离充足判据 [-] / Sufficient-distance verdict
    bStopRequest   : BOOL;             // 停车请求（MC_Halt 触发源）[-] / Stop request for MC_Halt
    bError         : BOOL;             // 故障锁存标志 [-] / Fault latch flag
    nErrId         : UDINT;            // 故障码，0 = 无故障（本件无信息码） / Fault code only
END_VAR
VAR
    _eState        : E_DL_AbpState := E_DL_AbpState.eIdle;   // 内部相位（CASE 唯一写入目标） / Internal phase
    _eCause        : E_DL_AbpCause := E_DL_AbpCause.eNone;   // 故障成因锁存（锁存量） / Latched cause
    rtReset        : R_TRIG;           // 复位沿实例，每周期无条件调用 / Reset edge
    _fReactMm      : REAL;             // 反应距离 [mm]（当拍量） / Reaction distance
    _fBrakeMm      : REAL;             // 制动距离 [mm]（当拍量） / Braking distance
    _fStopMm       : REAL;             // 停车总距离 [mm]（当拍量） / Total stopping distance
    _fAvailMm      : REAL;             // 可用距离 [mm]（当拍量） / Available distance
    _bStopOk       : BOOL;             // 判据（当拍量） / Verdict
    _bNonFin       : BOOL;             // 输入非有限当拍量 [-] / Non-finite input
    _bCfgBad       : BOOL;             // 组态非法当拍量 [-] / Config illegal
    _bFault        : BOOL;             // 故障锁存位（锁存量） / Latched fault bit
    _uFault        : UDINT;            // 故障码锁存（锁存量） / Latched fault code
END_VAR

(* —— 段 0：沿实例无条件周期刷新 + 当拍量判据（除零前置：减速度正域） —— *)
_bNonFin := (fActVelMmS <> fActVelMmS) OR (fPosMm <> fPosMm) OR (fLimitPosMm <> fLimitPosMm)
         OR ((fActVelMmS - fActVelMmS) <> (fActVelMmS - fActVelMmS))
         OR ((fPosMm - fPosMm) <> (fPosMm - fPosMm))
         OR ((fLimitPosMm - fLimitPosMm) <> (fLimitPosMm - fLimitPosMm));      // NaN 自反 + Inf 差值自减 / NaN and Inf
_bCfgBad := (fDecelMmS2 <= 1.0E-6) OR (tReaction <= T#0S) OR (fSafetyMarginMm < 0.0);   // 组态非法当拍量 / Config illegal
rtReset(CLK := bReset);                                                       // 复位沿，每拍必调 / Reset edge

(* —— 段 1：单拍量预清零（锁存量不入清单） —— *)
fStopDistMm := 0.0;                // 停车距离缺省 0 / Stopping distance default
fAvailMm := 0.0;                   // 可用距离缺省 0 / Available default
bStopOk := FALSE;                  // 判据缺省 FALSE（安全侧） / Verdict default safe
bStopRequest := TRUE;              // 停车请求缺省 TRUE（安全侧） / Stop request default safe
nErrId := 16#0000_0000;            // 故障码缺省无故障 / Fault code default

(* —— 段 2：复位沿 + 组态域闸 —— *)
IF rtReset.Q THEN                              // rtReset.Q = 当拍量 / current scan
    _bFault := FALSE;                          // 清故障锁存位（锁存量） / Clear fault latch
    _uFault := 16#0000_0000;                   // 清故障锁存码（锁存量） / Clear fault code
    _eCause := E_DL_AbpCause.eNone;            // 清成因（锁存量） / Clear cause
    IF _eState = E_DL_AbpState.eFault THEN
        _eState := E_DL_AbpState.eIdle;        // 故障相迁出：回未使能 / Fault exit to idle
    END_IF
END_IF
IF _bCfgBad THEN                               // 组态域闸 / Config gate
    _uFault := 16#0004_04A6;                   // 故障级：预判故障总码 / Motion fault code
    _eCause := E_DL_AbpCause.eCfgIllegal;      // 归因：组态非法 / Cause: illegal config
    _bFault := TRUE;                           // 标志与码位配对（R45） / Flag paired with code
END_IF
IF (NOT _bFault) AND _bNonFin THEN             // 非有限锁存 / Non-finite latch
    _uFault := 16#0004_04A6;
    _eCause := E_DL_AbpCause.eNonFinite;       // 归因：非有限 / Cause: non-finite
    _bFault := TRUE;
END_IF

(* —— 段 3：停车距离与可用距离计算（仅无故障；减速度已校验正域） —— *)
IF NOT _bFault THEN
    _fReactMm := fActVelMmS * (TIME_TO_REAL(tReaction) / 1000.0);              // 反应距离 [mm]（除常量 1000.0） / Reaction distance
    _fBrakeMm := fActVelMmS * fActVelMmS / (2.0 * fDecelMmS2);                 // 制动距离 [mm]（除数为已校验正域） / Braking distance
    _fStopMm := _fReactMm + _fBrakeMm + fSafetyMarginMm;                       // 停车总距离 [mm] / Total stopping distance
    IF bDirPositive THEN
        _fAvailMm := fLimitPosMm - fPosMm;                                     // 正向可用距离 / Positive available distance
    ELSE
        _fAvailMm := fPosMm - fLimitPosMm;                                     // 反向可用距离 / Negative available distance
    END_IF
    IF _fAvailMm < 0.0 THEN                                                    // 已越限位：可用距离钳制 0 / Clamp to zero
        _fAvailMm := 0.0;
    END_IF
    _bStopOk := _fAvailMm > _fStopMm;                                          // 判据（严格大于，含余量） / Verdict
END_IF

(* —— 段 4：故障解除式（R240；全当拍量）：rtReset.Q / NOT _bCfgBad / NOT _bNonFin —— *)
IF rtReset.Q AND (NOT _bCfgBad) AND (NOT _bNonFin) THEN
    _bFault := FALSE;                          // 清故障锁存位（锁存量） / Clear fault latch
    _uFault := 16#0000_0000;                   // 清故障锁存码（锁存量） / Clear fault code
    _eCause := E_DL_AbpCause.eNone;            // 清成因（锁存量） / Clear cause
END_IF

(* —— 段 4A：故障锁存相位迁移闸（请求停车） —— *)
IF _bFault AND (_eState <> E_DL_AbpState.eFault) THEN
    _eState := E_DL_AbpState.eFault;           // 锁存即入故障相 / Latch enters fault phase
END_IF

(* —— 段 5：相位机（CASE 全覆盖 + ELSE 兜底） —— *)
CASE _eState OF

E_DL_AbpState.eIdle:
    IF bEnable AND (NOT _bFault) THEN          // 使能条件 / Enable gate
        _eState := E_DL_AbpState.eRun;         // 进预判相 / Enter prediction
    END_IF

E_DL_AbpState.eRun:
    IF NOT _bStopOk THEN                       // 出口 1：距离不足（事件） / Insufficient distance
        _eState := E_DL_AbpState.eBrake;       // 进请求停车相 / Enter stop request
    ELSIF NOT bEnable THEN                     // 出口 2：撤使能（前置消失） / Disable
        _eState := E_DL_AbpState.eIdle;
    END_IF

E_DL_AbpState.eBrake:
    IF _bStopOk AND bEnable THEN               // 距离恢复充足：回预判相 / Distance sufficient again
        _eState := E_DL_AbpState.eRun;
    ELSIF NOT bEnable THEN                     // 撤使能：回未使能 / Disable returns idle
        _eState := E_DL_AbpState.eIdle;
    END_IF

E_DL_AbpState.eFault:
    ;                                          // 故障相：请求停车，仅段 4 复位沿可迁出 / Stop requested, reset only

ELSE
    _uFault := 16#0004_04A6;                   // 故障级：非法相位兜底（归并总码） / Illegal phase fallback
    _eCause := E_DL_AbpCause.eCfgIllegal;      // 归因：相位非法归并组态 / Cause: phase illegal
    _bFault := TRUE;
    _eState := E_DL_AbpState.eFault;           // 强制回故障相 / Force fault phase

END_CASE

(* —— 段 6：出口单点映射（名实同源；故障相请求停车） —— *)
IF _bFault THEN
    nErrId := _uFault;                         // 故障锁存码回放 / Replay latched code
    bStopOk := FALSE;                          // 故障相判据强制 FALSE（安全侧） / Verdict forced false
    bStopRequest := TRUE;                      // 故障相请求停车 / Stop requested
    fStopDistMm := 0.0;                        // 故障相距离出口强制 0 / Distance forced zero
    fAvailMm := 0.0;                           // 故障相可用距离强制 0 / Available forced zero
ELSE
    nErrId := 16#0000_0000;                    // 无故障：本件无信息码 / No fault, no info code
    bStopOk := _bStopOk;                       // 判据出口 / Verdict outlet
    bStopRequest := (_eState = E_DL_AbpState.eBrake) OR (NOT _bStopOk);   // 停车请求出口 / Stop request outlet
    fStopDistMm := _fStopMm;                   // 停车距离出口 / Distance outlet
    fAvailMm := _fAvailMm;                     // 可用距离出口 / Available outlet
END_IF
bError := _bFault;                             // 故障标志同源 / Flag from latch
eState := _eState;                             // 状态出口 / State outlet
eCause := _eCause;                             // 成因出口 / Cause outlet

END_FUNCTION_BLOCK

(* ---- FB_DL_AxisBrakeTest.st ---- *)
(*
  组件名 Component   : FB_DL_AxisBrakeTest
  子库 Sublibrary    : DL_Motion
  版本 Version       : 1.0.0
  兼容性 Platform    : CODESYS 3.5 / TwinCAT 3 / 汇川 InoProShop / Machine Expert（仅 Standard.library）
  功能 Function      : 抱闸制动测试顺控（与 FB_DL_AxisBrakeDistPredict 分工：预测制动
                       距离 vs 周期性制动测试）：
                       1) 测试以上升沿承载：eIdle → eCloseBrake（出抱闸闭合指令）；
                       2) eCloseBrake：等轴零速（|速度| < 近零阈 持续 tZeroWin 确认），
                       超时 tZeroTo 判故障；抱闸反馈缺失判故障；
                       3) eMeasure：位置快照后驻留 tHoldDur，滑移量 = |位置 - 快照|，
                       超过 fSlipLimitMm 判不合格，否则合格；
                       4) eDone：结果驻留至测试指令撤销；到期计数按使能期扫描累计，
                       超过 uTestIntervalScans 置 bTestDue。
  边界 Boundary      : ① 本件只出抱闸闭合指令与测试结论，不驱动运动指令；
                       ② 各相超时用独立 TON 实例（tonZeroTo / tonHoldDur），禁跨相复用；
                       ③ 滑移量除法无（纯差值比较），非有限输入判非法锁存；
                       ④ 故障锁存解除唯一路径 = bReset 上升沿（输入引脚，恒可达）；
                       ⑤ 无全局变量引用、无外部变量声明、无物理地址寻址。
  依赖 Depends       : Standard.library（R_TRIG / TON）
  溯源 Origin        : 道莅自研 clean-room（参考 t1-6-plcopen 运动接口分类与参数域，
                       零代码行复制）
  码位 Code          : 16#04_0_AA
  码表 Error codes（Motion 格 04_0_AA，单轨：故障 0x02AA / 信息 0x01AA）:
    16#0004_02AA 故障级：测试非法（零速超时 / 抱闸反馈缺失 / 组态非法 / 输入非有限），
                 锁存至 bReset 上升沿
    16#0004_01AA 信息级：测试结论写定沿（合格或不合格判定拍，bTestPass 同拍定值）
  修订历史 Revision  :
    2026-11-19  v1.0.0  R44 首版（批次 2 · 序号 7）
*)

TYPE E_DL_AbtState :
(
    eIdle       := 0,   // 空闲：等测试沿 / Idle, waiting test edge
    eCloseBrake := 10,  // 闭闸：等零速确认 / Closing brake, waiting zero speed
    eMeasure    := 20,  // 测量：驻留计滑移 / Measuring, slip dwell
    eDone       := 30,  // 完成：结论驻留 / Done, verdict held
    eFault      := 90   // 故障：测试非法锁存 / Fault, latched
);
END_TYPE

FUNCTION_BLOCK FB_DL_AxisBrakeTest
VAR_INPUT
    bEnable        : BOOL;               // 使能（电平），使能期累计到期计数 [-] / Enable
    bReset         : BOOL;               // 上升沿清故障锁存 [-] / Reset edge
    bTestCmd       : BOOL;               // 测试指令（上升沿承载）[-] / Test command edge
    fVelMmS        : REAL;               // 轴实际速度 [mm/s] / Axis velocity
    fPosMm         : REAL;               // 轴实际位置 [mm] / Axis position
    bBrakeFb       : BOOL;               // 抱闸闭合反馈 [-] / Brake closed feedback
    fVelNearZeroMmS: REAL := 0.5;        // 零速判据阈 [mm/s] / Near-zero velocity threshold
    fSlipLimitMm   : REAL := 0.1;        // 滑移量合格限 [mm] / Slip pass limit
    tZeroWin       : TIME := T#500MS;    // 零速确认窗 [毫秒] / Zero-speed confirm window
    tZeroTo        : TIME := T#10S;      // 闭闸零速超时 [毫秒] / Zero-speed timeout
    tHoldDur       : TIME := T#5S;       // 滑移测量驻留 [毫秒] / Slip measurement dwell
    uTestIntervalScans: UDINT := 8640000;// 定期测试到期计数 [拍] / Test due interval in scans
END_VAR
VAR_OUTPUT
    bBrakeCmdOut   : BOOL;               // 抱闸闭合指令输出 [-] / Brake close command
    bTestBusy      : BOOL;               // 测试进行中电平 [-] / Test busy level
    bTestPass      : BOOL;               // 结论：TRUE = 合格 [-] / Verdict pass flag
    bTestDue       : BOOL;               // 定期测试到期标志 [-] / Test due flag
    fSlipMm        : REAL;               // 实测滑移量 [mm] / Measured slip
    uScansSinceTest: UDINT;              // 距上次测试扫描累计 [拍] / Scans since last test
    eState         : E_DL_AbtState;      // 状态出口，段尾单点映射 / State outlet
    bError         : BOOL;               // 故障锁存标志 [-] / Fault latch flag
    uErrId         : UDINT;              // 事件码，0 = 无事件 / Event code
END_VAR
VAR
    rtReset  : R_TRIG;                   // 复位沿实例，段 0 无条件刷新 / Reset edge
    rtTest   : R_TRIG;                   // 测试沿实例，段 0 无条件刷新 / Test edge
    tonZeroWin: TON;                     // 零速确认窗 / Zero-speed confirm timer
    tonZeroTo : TON;                     // 闭闸超时（专用超时件命名） / Zero-speed timeout
    tonHoldDur: TON;                     // 测量驻留计时 / Measurement dwell timer
    _eState  : E_DL_AbtState := E_DL_AbtState.eIdle;   // 内部相位（CASE 唯一写入目标）/ Internal phase
    _fPosSnap: REAL;                     // 测量起点位置快照 [mm] / Position snapshot
    _bFault  : BOOL;                     // 故障锁存位（锁存量） / Latched fault bit
    _uFault  : UDINT;                    // 故障码锁存（锁存量） / Latched fault code
    _bCfgBad : BOOL;                     // 组态非法当拍量 [-] / Config illegal flag
    _bNonFin : BOOL;                     // 输入非有限当拍量 [-] / Non-finite input flag
END_VAR
VAR CONSTANT
    DL_ABS_MAX : REAL := 1.0E30;         // 有限值判定上界 [工程单位] / Finite bound
    DL_ZERO    : REAL := 0.0;            // 零常量 [mm] / Zero constant
END_VAR

(* —— 段 0｜沿与定时器每拍无条件刷新（禁置于 IF/CASE 内） —— *)
rtReset(CLK := bReset);
rtTest (CLK := bTestCmd);
tonZeroWin (IN := (_eState = E_DL_AbtState.eCloseBrake) AND (ABS(fVelMmS) < fVelNearZeroMmS)
             AND (NOT _bFault), PT := tZeroWin);
tonZeroTo  (IN := (_eState = E_DL_AbtState.eCloseBrake) AND (NOT _bFault), PT := tZeroTo);
tonHoldDur (IN := (_eState = E_DL_AbtState.eMeasure) AND (NOT _bFault), PT := tHoldDur);

(* —— 段 1｜瞬时量预清零（锁存量 _bFault/_uFault/bTestPass/_fPosSnap 不入清单） —— *)
uErrId   := 16#0000_0000;
_bCfgBad := FALSE;
_bNonFin := FALSE;

(* —— 段 2｜复位沿：故障一次性清干净，相位回空闲，抱闸指令撤销 —— *)
IF rtReset.Q THEN
    _bFault  := FALSE;
    _uFault  := 16#0000_0000;
    bBrakeCmdOut := FALSE;
    _eState  := E_DL_AbtState.eIdle;
END_IF

(* —— 段 3｜组态闸与非有限判据 —— *)
IF (fVelNearZeroMmS <= DL_ZERO) OR (fSlipLimitMm <= DL_ZERO) OR (tZeroWin = T#0S)
   OR (tZeroTo = T#0S) OR (tHoldDur = T#0S) THEN
    _bCfgBad := TRUE;
END_IF
IF (fVelMmS <> fVelMmS) OR ((fVelMmS - fVelMmS) <> DL_ZERO)
   OR (fPosMm <> fPosMm) OR ((fPosMm - fPosMm) <> DL_ZERO) THEN
    _bNonFin := TRUE;
END_IF

(* —— 段 4｜到期计数：使能期每拍累计，超限置到期标志 —— *)
IF bEnable AND (NOT _bFault) THEN
    uScansSinceTest := uScansSinceTest + UDINT#1;
    IF uScansSinceTest >= uTestIntervalScans THEN
        bTestDue := TRUE;
    END_IF
END_IF

(* —— 段 5｜主状态机：五态全覆盖 + ELSE 兜底 —— *)
CASE _eState OF

E_DL_AbtState.eIdle:
    bBrakeCmdOut := FALSE;
    bTestBusy    := FALSE;
    IF _bFault THEN
        bError := TRUE;                  // 故障锁存回放（R189）
    END_IF
    IF rtTest.Q AND bEnable AND (NOT _bFault) AND (NOT _bCfgBad) AND (NOT _bNonFin) THEN
        uScansSinceTest := UDINT#0;      // 新测试起点：到期计数清零
        bTestDue := FALSE;
        bBrakeCmdOut := TRUE;            // 出抱闸闭合指令
        bTestBusy := TRUE;
        _eState := E_DL_AbtState.eCloseBrake;
    ELSIF rtTest.Q AND (_bCfgBad OR _bNonFin OR _bFault) THEN
        _bFault := TRUE;                 // 带病启动拒绝
        _uFault := 16#0004_02AA;
        bError  := TRUE;
        _eState := E_DL_AbtState.eFault;
    END_IF

E_DL_AbtState.eCloseBrake:
    bBrakeCmdOut := TRUE;
    bTestBusy := TRUE;
    IF _bNonFin THEN
        _bFault := TRUE;                 // 输入非有限：判据不可信
        _uFault := 16#0004_02AA;
        bError  := TRUE;
        _eState := E_DL_AbtState.eFault;
    ELSIF NOT bBrakeFb THEN
        _bFault := TRUE;                 // 抱闸反馈缺失：指令已出而反馈不到
        _uFault := 16#0004_02AA;
        bError  := TRUE;
        _eState := E_DL_AbtState.eFault;
    ELSIF tonZeroWin.Q THEN
        _fPosSnap := fPosMm;             // 零速确认：取滑移测量起点快照
        _eState := E_DL_AbtState.eMeasure;   // 迁出条件 1：零速达成
    ELSIF tonZeroTo.Q THEN
        _bFault := TRUE;                 // 迁出条件 2（故障路）：零速超时
        _uFault := 16#0004_02AA;
        bError  := TRUE;
        _eState := E_DL_AbtState.eFault;
    END_IF

E_DL_AbtState.eMeasure:
    bBrakeCmdOut := TRUE;
    bTestBusy := TRUE;
    IF tonHoldDur.Q THEN
        fSlipMm := ABS(fPosMm - _fPosSnap);  // 滑移量 = 驻留期位置漂移
        bTestPass := fSlipMm <= fSlipLimitMm;
        uErrId := 16#0004_01AA;          // 信息级：结论写定沿（锁存至复位）
        _eState := E_DL_AbtState.eDone;
    END_IF

E_DL_AbtState.eDone:
    bBrakeCmdOut := FALSE;               // 测试结束：抱闸指令撤销
    bTestBusy := FALSE;
    IF NOT bTestCmd THEN
        _eState := E_DL_AbtState.eIdle;  // 测试指令撤销：回空闲（结论锁存保留）
    END_IF

E_DL_AbtState.eFault:
    bBrakeCmdOut := FALSE;               // 故障相：抱闸指令安全侧撤销
    bTestBusy := FALSE;
    bError := TRUE;
    ;                                    // 故障相驻留：只认复位沿（段 2 迁出）

ELSE
    _bFault := TRUE;                     // 兜底：非法相位锁存
    _uFault := 16#0004_02AA;
    bError  := TRUE;
    _eState := E_DL_AbtState.eFault;
END_CASE

(* —— 段 6｜状态出口单点映射 —— *)
eState := _eState;
END_FUNCTION_BLOCK

(* ---- FB_DL_AxisCantileverComp.st ---- *)
(*
  ==================================================================
  组件名 Component  : FB_DL_AxisCantileverComp
  分类   Category   : DL_Motion
  复杂度 Complexity  : cx4
  版本   Version    : 1.0.0
  功能   Purpose    : 悬臂轴重力下垂补偿。按位置 pos 在段点表（afSegX / afSegC，
                      基准负载下的补偿曲线）分段线性插值，再按实际负载与基准负载
                      之比缩放，得补偿量 fComp 叠加到位置指令；补偿上限钳制；
                      负载超上限判 ePayloadOver；曲表段点不严格递增判
                      eCurveDegenerate；上电首拍不输出补偿（自零起斜坡引入，
                      单拍步进上限 fStepMax）。
  来源   Source     : t1-6-plcopen（limits / comp 族）
  溯源   Origin     : IEC 61131-3 标准语义的道莅防御性实现；悬臂挠曲随负载 / 伸长
                      量的材料力学前馈修正为公开力学语义，clean-room 自研实现，
                      未复制任何闭源代码行。
  平台   Platform   : 纯 IEC 61131-3（ARRAY / LREAL 运算，无私有库、无幂运算符）
  作者   Author     : 道莅代码库 · PLC 编程专家（R56）
  ------------------------------------------------------------------
  边界 Boundary     :
                      一 本件只算补偿量，不驱动轴、不改位置环（属主边界）；
                      二 故障优先级固定：eSensorBad > eCurveDegenerate > ePayloadOver
                         （R146 方向性：传感器失效冻结，曲表失效不输出，负载超限降级钳制）；
                      三 首拍斜坡：出口自零起按 fStepMax 单拍步进逼近目标（首拍不跳变）；
                      四 故障锁存（曲表退化 / 负载超限）解除路径 = bReset 上升沿（R188）；
                      五 无全局变量、无外部变量声明、无物理地址寻址。
  输出契约 Output contract:
                      fComp 为斜坡后的补偿量出口 [位置单位]；
                      eFault 为锁存回放；ePhaseBad 为非法相位兜底专用成员（R128）。
  修订记录 Revision  :
    2026-11-20  v1.0.0  R56 首版（批 3 · 序号 13）
  ==================================================================
*)

TYPE E_DL_AcfPhase :
(
    eIdle  := 0,  // 未使能：出口保持 / disabled, the outlet holds
    eRun   := 10, // 运行：逐拍插值与斜坡 / running, interpolation and the ramp every scan
    eFault := 90  // 故障：成因锁存，出口冻结 / fault, the cause is latched, the outlet freezes
);
END_TYPE

TYPE E_DL_AcfFault :
(
    eNone             := 0, // 无成因 / no cause
    eCurveDegenerate  := 1, // 曲表退化：段点不严格递增或段数不足（故障级，与 bError 配对）/ a degenerate curve, fault grade paired with bError
    ePayloadOver      := 2, // 负载超上限（信息级，补偿按上限钳制）/ the payload is over the ceiling, the compensation clamps
    eSensorBad        := 3, // 位置或负载非有限（故障级，与 bError 配对）/ the position or the load is non finite, fault grade paired with bError
    ePhaseBad         := 4  // 非法相位兜底（故障级，与 bError 配对）/ illegal phase fallback, fault grade paired with bError
);
END_TYPE

FUNCTION_BLOCK FB_DL_AxisCantileverComp
VAR_INPUT
    bEnable  : BOOL := TRUE;    // 使能，失能时出口冻结保持 [-] / enable, the outlet holds when disabled
    bReset   : BOOL := FALSE;   // 复位上升沿清故障锁存并出口归零 [-] / reset rising edge clears the latch and zeroes the outlet
    fPos     : LREAL := 0.0;    // 轴实际位置 [位置单位] / the actual axis position [position unit]
    fLoadKg  : LREAL := 0.0;    // 负载质量 [千克] / the payload mass [kilogram]
    fLoadRef : LREAL := 10.0;   // 曲表基准负载 [千克]，域 大于零 / the curve reference load [kilogram], domain above zero
    fLoadMax : LREAL := 50.0;   // 负载上限 [千克]，域 大于零 / the payload ceiling [kilogram], domain above zero
    fCompMax : LREAL := 1.0;    // 补偿量上限 [位置单位]，域 大于零 / the compensation ceiling [position unit], domain above zero
    fStepMax : LREAL := 0.01;   // 首拍斜坡单拍步进上限 [位置单位每拍]，0 = 直通 / the ramp step ceiling per scan, zero is a passthrough
    afSegX   : ARRAY[1..16] OF LREAL := [0.0, 100.0, 200.0, 300.0, 400.0, 500.0, 600.0, 700.0, 800.0, 900.0, 1000.0, 0.0, 0.0, 0.0, 0.0, 0.0]; // 段点位置表（升序有效段）[位置单位] / the segment position table in ascending order [position unit]
    afSegC   : ARRAY[1..16] OF LREAL := [16(0.0)]; // 段点补偿量表（基准负载下）[位置单位] / the segment compensation table at the reference load [position unit]
    nSeg     : INT := 11;       // 有效段点数 [个]，域 2..16 / the valid segment count, domain two to sixteen
END_VAR
VAR_OUTPUT
    fComp    : LREAL := 0.0;  // 补偿量出口（叠加到位置指令）[位置单位] / the compensation outlet for the position command [position unit]
    ePhase   : E_DL_AcfPhase := E_DL_AcfPhase.eIdle; // 相位出口 [枚举] / phase outlet [enum]
    eFault   : E_DL_AcfFault := E_DL_AcfFault.eNone; // 成因出口，锁存回放 [枚举] / cause outlet replayed from the latch [enum]
    bError   : BOOL := FALSE; // 故障锁存标志 [-] / fault latch flag
END_VAR
VAR
    rtReset  : R_TRIG; // 复位沿检测，段 0 无条件刷新 / reset edge, refreshed unconditionally in segment zero
    _ePhase  : E_DL_AcfPhase := E_DL_AcfPhase.eIdle; // 内部相位，CASE 唯一写入目标 / internal phase, the only CASE write target
    _eFaulC  : E_DL_AcfFault := E_DL_AcfFault.eNone; // 故障级成因，锁存至复位沿 / fault cause, latched until the reset edge
    _bFault  : BOOL := FALSE; // 故障锁存位 [-] / fault latch bit
    _bInit   : BOOL := FALSE; // 首扫初始化完成标志（R310）/ first scan initialisation flag
    _bInOk   : BOOL := FALSE; // 位置与负载均有限 [-] / both position and load are finite
    _bCfgOk  : BOOL := FALSE; // 组态参数域内 [-] / the configuration is inside the domain
    _bCurveOk: BOOL := FALSE; // 曲表结构合法 [-] / the curve structure is legal
    _bPayload: BOOL := FALSE; // 负载超上限标志 [-] / the payload over ceiling flag
    _nSegUse : INT := 11;     // 钳定后的段点数 [个] / the clamped segment count
    _nI      : INT := 1;      // 插值段游标 [段] / the interpolation segment cursor
    _nGuard  : INT := 0;      // 扫描守护计数 [次] / the scan guard [count]
    _fScale  : LREAL := 1.0;  // 负载缩放比 [无量纲] / the load scale ratio
    _fLoadUse: LREAL := 0.0;  // 钳定后的负载 [千克] / the clamped load [kilogram]
    _fTarget : LREAL := 0.0;  // 本拍补偿目标值 [位置单位] / the compensation target this scan [position unit]
    _fStep   : LREAL := 0.0;  // 本拍步进量 [位置单位] / the step this scan [position unit]
END_VAR

// 段 0｜沿检测无条件周期刷新（禁入分支）/ segment 0, unconditional refresh of the edge detector
rtReset(CLK := bReset); // 复位沿无条件刷新 / unconditional refresh of the reset edge

// 段 1｜首扫初始化（R310）：出口自零起步（首拍不输出补偿）/ segment 1, first scan initialisation, the outlet starts at zero
IF NOT _bInit THEN // 首扫一拍 / the very first scan
    _bInit := TRUE; // 置首扫完成标志 / raise the first scan flag
    _ePhase := E_DL_AcfPhase.eRun; // 相位从运行起步 / the phase starts in run
    _eFaulC := E_DL_AcfFault.eNone; // 故障级成因清零 / clear the fault cause
    _bFault := FALSE; // 故障锁存清零 / clear the fault latch
    fComp := 0.0; // 出口自零起步（首拍斜坡引入）/ the outlet starts at zero for the ramp in
END_IF

// 段 2｜复位沿作用域：清锁存 / 迁相位 / 出口归零（三项逐项声明）/ segment 2, reset edge scope declared item by item
IF rtReset.Q THEN // 复位沿 / the reset edge
    _bFault := FALSE; // 作用域一：清故障锁存 / scope one, clear the fault latch
    _eFaulC := E_DL_AcfFault.eNone; // 作用域一：清故障级成因 / scope one, clear the fault cause
    _ePhase := E_DL_AcfPhase.eRun; // 作用域二：迁回运行相 / scope two, migrate back to run
    fComp := 0.0; // 作用域三：出口归零（斜坡自零重引入）/ scope three, the outlet zeroes for a fresh ramp
END_IF

// 段 3｜组态域闸与曲表结构校验（R151 全覆盖）/ segment 3, the configuration gate and the curve structure check
_bInOk := (fPos = fPos) AND ((fPos - fPos) = (fPos - fPos)) AND (fLoadKg = fLoadKg) AND ((fLoadKg - fLoadKg) = (fLoadKg - fLoadKg)); // 位置与负载有限性 / finiteness of the position and the load
_bCfgOk := (fLoadRef > 0.0) AND (fLoadRef = fLoadRef) AND (fLoadMax > 0.0) AND (fLoadMax = fLoadMax) AND (fCompMax > 0.0) AND (fCompMax = fCompMax) AND (fStepMax >= 0.0) AND (fStepMax = fStepMax); // 组态参数域判定 / the configuration domain verdict
_nSegUse := nSeg; // 段点数直通 / the segment count passes through
IF _nSegUse < 2 THEN // 下越域 / below the floor
    _nSegUse := 2; // 回钳到二 / clamp to two
ELSIF _nSegUse > 16 THEN // 上越域 / above the ceiling
    _nSegUse := 16; // 回钳到十六 / clamp to sixteen
END_IF
_bCurveOk := _bCfgOk AND (_nSegUse >= 2); // 曲表结构初判 / the first curve verdict
_nI := 1; // 扫描游标起步 / start the scan cursor
_nGuard := 0; // 守护清零 / clear the guard
WHILE (_nI < _nSegUse) AND (_nGuard < 16) DO // 严格递增校验，守护为容量 / the strict monotonic check with the capacity as the guard
    _nGuard := _nGuard + 1; // 守护递增 / increment the guard
    IF afSegX[_nI] >= afSegX[_nI + 1] THEN // 段点非严格递增 / the points are not strictly increasing
        _bCurveOk := FALSE; // 判曲表退化 / the curve is degenerate
    END_IF
    _nI := _nI + 1; // 游标递增 / increment the cursor
END_WHILE

// 段 4｜相位机：ENUM + CASE，含 ELSE 非法相位兜底（R128）/ segment 4, the phase machine with an ELSE fallback
CASE _ePhase OF
E_DL_AcfPhase.eIdle: // 未使能相：出口冻结保持 / the disabled phase, the outlet holds
    IF bEnable AND (NOT _bFault) THEN // 使能且无故障 / enabled and unfaulted
        _ePhase := E_DL_AcfPhase.eRun; // 迁运行相 / migrate to run
    END_IF

E_DL_AcfPhase.eRun: // 运行相：插值 + 缩放 + 钳制 + 斜坡 / the run phase, interpolate, scale, clamp and ramp
    IF NOT bEnable THEN // 失能 / disabled
        _ePhase := E_DL_AcfPhase.eIdle; // 迁未使能相 / migrate to idle
    ELSIF (NOT _bInOk) OR (NOT _bCurveOk) THEN // 传感器失效或曲表退化（高优先级拦截）/ a sensor failure or a degenerate curve, the top priority interception
        _bFault := TRUE; // 置故障锁存 / raise the fault latch
        IF NOT _bInOk THEN // 传感器失效优先归因（R190 独立成因）/ the sensor failure takes the cause priority
            _eFaulC := E_DL_AcfFault.eSensorBad; // 故障级成因（R45 配对 bError）/ the fault cause paired with bError
        ELSE // 曲表退化归因 / the degenerate curve cause
            _eFaulC := E_DL_AcfFault.eCurveDegenerate; // 故障级成因（R45 配对 bError）/ the fault cause paired with bError
        END_IF
        _ePhase := E_DL_AcfPhase.eFault; // 迁故障相 / migrate to the fault phase
    ELSE // 正常计算 / the normal computation
        _fLoadUse := fLoadKg; // 负载直通 / the load passes through
        _bPayload := FALSE; // 负载超限标志预置假 / preset the payload flag to false
        IF _fLoadUse < 0.0 THEN // 负载负值回钳零 / a negative load clamps to zero
            _fLoadUse := 0.0; // 钳到零 / clamp to zero
        ELSIF _fLoadUse > fLoadMax THEN // 负载超上限 / the load is over the ceiling
            _fLoadUse := fLoadMax; // 钳到上限（信息级降级，R146 安全侧）/ clamp to the ceiling, the safe side
            _bPayload := TRUE; // 置负载超限标志 / raise the payload flag
        END_IF
        _fScale := _fLoadUse / fLoadRef; // 负载缩放比，除子为基准负载已证大于零 / the load scale with the proven reference divisor
        _fTarget := 0.0; // 目标值预置零 / preset the target to zero
        IF fPos <= afSegX[1] THEN // 左端外推钳位 / below the first point
            _fTarget := afSegC[1] * _fScale; // 取首段点补偿 / take the first point compensation
        ELSIF fPos >= afSegX[_nSegUse] THEN // 右端外推钳位 / above the last point
            _fTarget := afSegC[_nSegUse] * _fScale; // 取末段点补偿 / take the last point compensation
        ELSE // 域内分段线性插值 / the in domain piecewise interpolation
            _nI := 1; // 段游标起步 / start the segment cursor
            _nGuard := 0; // 守护清零 / clear the guard
            WHILE (_nI < _nSegUse) AND (_nGuard < 16) AND (fPos > afSegX[_nI + 1]) DO // 定位所在段 / locate the segment
                _nGuard := _nGuard + 1; // 守护递增 / increment the guard
                _nI := _nI + 1; // 游标递增 / increment the cursor
            END_WHILE
            _fTarget := afSegC[_nI] + (afSegC[_nI + 1] - afSegC[_nI]) * (fPos - afSegX[_nI]) / (afSegX[_nI + 1] - afSegX[_nI]); // 线性插值，除子为段宽已证大于零（严格递增校验）/ the linear interpolation with the proven segment width
            _fTarget := _fTarget * _fScale; // 负载缩放 / scale by the load
        END_IF
        IF _fTarget > fCompMax THEN // 补偿上限钳制 / clamp the compensation high
            _fTarget := fCompMax; // 钳到上限 / clamp to the ceiling
        ELSIF _fTarget < -fCompMax THEN // 补偿下限钳制 / clamp the compensation low
            _fTarget := -fCompMax; // 钳到下限 / clamp to the floor
        END_IF
        IF fStepMax <= 0.0 THEN // 步进上限为零 = 直通 / a zero step means a passthrough
            fComp := _fTarget; // 直通出口 / the passthrough outlet
        ELSE // 斜坡逼近 / the ramp approach
            _fStep := _fTarget - fComp; // 本拍剩余差 / the remaining difference
            IF _fStep > fStepMax THEN // 上行限步 / limit the upward step
                _fStep := fStepMax; // 钳到步进上限 / clamp to the step ceiling
            ELSIF _fStep < -fStepMax THEN // 下行限步 / limit the downward step
                _fStep := -fStepMax; // 钳到步进下限 / clamp to the step floor
            END_IF
            fComp := fComp + _fStep; // 斜坡推进 / advance the ramp
        END_IF
        IF _bPayload THEN // 负载超限信息级（不置故障锁存，R146 降级方向）/ the payload flag is informational, a degrade direction
            _eFaulC := E_DL_AcfFault.ePayloadOver; // 信息级成因 / the informational cause
        ELSE // 恢复后撤销 / revoked on recovery
            _eFaulC := E_DL_AcfFault.eNone; // 成因清零 / clear the cause
        END_IF
    END_IF

E_DL_AcfPhase.eFault: // 故障相：出口冻结保持，等复位沿 / the fault phase, the outlet freezes until the reset edge
    IF NOT bEnable THEN // 失能 / disabled
        _ePhase := E_DL_AcfPhase.eIdle; // 迁未使能相 / migrate to idle
    END_IF

ELSE // 非法相位兜底（R128）/ the illegal phase fallback
    _bFault := TRUE; // 置故障锁存 / raise the fault latch
    _eFaulC := E_DL_AcfFault.ePhaseBad; // 故障级成因（R45 配对 bError）/ the fault cause paired with bError
    _ePhase := E_DL_AcfPhase.eFault; // 迁故障相 / migrate to the fault phase
END_CASE

// 段 5｜统一出口 / segment 5, the unified outlet
IF _bFault THEN // 故障锁存优先 / the fault latch takes priority
    eFault := _eFaulC; // 故障级成因锁存回放（R152）/ the fault cause replayed from the latch
ELSE
    eFault := _eFaulC; // 信息级成因直映 / the informational cause is mapped directly
END_IF
ePhase := _ePhase; // 相位出口单点映射 / single point phase outlet mapping
bError := _bFault; // 故障标志与锁存位同源 / the fault flag shares the latch source
END_FUNCTION_BLOCK

(* ---- FB_DL_AxisCmdArbiter.st ---- *)
(*
  ==================================================================
  组件名 Component  : FB_DL_AxisCmdArbiter
  分类   Category   : DL_Motion
  复杂度 Complexity  : 中
  版本   Version    : 1.0.1
  功能   Purpose    : 轴驱动命令源优先级仲裁。四级命令源 安全 > 手动 > 自动 > 上位，
                      每拍全量重判，输出胜出源标签与整份命令字（携带源身份，
                      防「赢了仲裁丢了身份」），源切换出单拍脉冲。
  来源   Source     : t1-6-plcopen（PLCopen 运动接口命令源语义）
  溯源   Origin     : 命令源优先级仲裁属公开运动控制语义，clean-room 自研实现，
                      未复制 PLCopen 官方库或任何厂商源码。
  平台   Platform   : 纯 IEC 61131-3（IF / ELSIF / CASE / 标准转换函数），三平台通用
  分工声明 Split     : 与 FB_DL_ModeArbiter（单元模式级属主）分工——后者仲裁整机/
                      单元运行模式；本件只仲裁单轴驱动命令源，不发运动指令、
                      不判轴状态、不自造轴状态枚举（PLCopen 纪律，R277）。
  作者   Author     : 道莅代码库 · PLC 编程专家（R60）
  ------------------------------------------------------------------
  归属 Ownership     : E_DL_AxisCmdSrc 与 ST_DL_AxisCmd 的属主为本文件（全库唯一
                      定义，R264）；引用件只引用不重声明。
  边界 Boundary     :
                      一 纯组合件，每拍全量重判，无相位机（R227 显式声明）：不存在
                         等待相、不存在陈旧保持，胜出结果即本拍输入的函数；
                      二 优先级写死 安全(10) > 手动(20) > 自动(30) > 上位(40)，
                         枚举数值小者优先；源标签不符（如 stSafe 携带 eAuto）
                         视为该源未请求，不参与仲裁；
                      三 输出命令字整体取自胜出源结构体并回写胜出源标签，调用方
                         据 eWinner 与 stWinnerCmd.eSrc 双重可判来源；
                      四 源切换单拍脉冲 bSwitched 统一出口段每拍先预置 FALSE、
                         分支只写 TRUE（R256）；
                      五 无请求源时输出 eNone 与安全侧零命令（bAnyActive = FALSE）；
                      六 使能 bEnable = FALSE 时语义为「降级为零命令 + 置标志」
                         （eWinner = eNone），不保持上拍命令（R191 声明行）；
                      七 有界豁免登记（R272，D11 返修）：非有限闸只判胜出源 _stWin
                         的两个浮点字段——非胜出源命令字不入出口、不参与判据
                         换算，属有界豁免（机检口径 2/8 显式声明，非漏闸）。
  错误码   Codes    :
    16#0004_0620【信息级】本拍无任何命令源请求（胜出 eNone）
    16#0004_0621【信息级】发生源切换（bSwitched 同拍置位）
    16#0004_0622【故障级】胜出源命令字含非有限量，已降级为零命令
  验收   Acceptance :
    算法已证（脚本）：未跑 ｜ 编译器已证（三平台）：未跑
    V1 仅自动源请求 → eWinner = eAuto、命令字等于自动源
    V2 安全源与手动源同拍请求 → eWinner = eSafe（小者优先）
    V3 全部源 eNone → eWinner = eNone、命令零值、码 0620
  修订记录 Revision  :
    2026-11-21  v1.0.0  R60 首版（批 3 · 序号 11）
    2026-11-21  v1.0.1  R61 返修：D1 降级路径 _eWinner 同步落 eNone（双通道
                        一致）；D2 增 _bFault 锁存位 + bReset 复位引脚，bError
                        改为锁存回放口径（R187）；D11 边界段登记非胜出源豁免
  ==================================================================
*)

TYPE E_DL_AxisCmdSrc :
(
    eNone := 0,  // 无源：本拍无命令请求 / none, no command source requests this scan
    eSafe := 10, // 安全源：最高优先级 / the safety source with the top priority
    eJog  := 20, // 手动源：次高优先级 / the jog source
    eAuto := 30, // 自动源：第三优先级 / the automatic source
    eHost := 40  // 上位源：最低优先级 / the host source with the lowest priority
);
END_TYPE

TYPE ST_DL_AxisCmd :
STRUCT
    eSrc     : E_DL_AxisCmdSrc := E_DL_AxisCmdSrc.eNone; // 命令来源标签 [源] / the command source label
    fVelMmS  : LREAL := 0.0;                             // 速度指令 [毫米每秒] / the velocity command
    fPosMm   : LREAL := 0.0;                             // 位置指令 [毫米] / the position command
    uFlags   : UDINT := 16#0000_0000;                    // 命令标志位 [位图] / the command flag word
END_STRUCT
END_TYPE

FUNCTION_BLOCK FB_DL_AxisCmdArbiter
VAR_INPUT
    bEnable : BOOL := TRUE;              // 使能，FALSE 时降级为零命令（边界六）/ the enable, false degrades to the zero command
    bReset  : BOOL := FALSE;             // 故障复位电平，上升沿清非有限故障锁存（D2 返修新增）/ the fault reset level, the rising edge clears the non finite latch
    stSafe  : ST_DL_AxisCmd;             // 安全源命令字 [源结构] / the safety source command
    stJog   : ST_DL_AxisCmd;             // 手动源命令字 [源结构] / the jog source command
    stAuto  : ST_DL_AxisCmd;             // 自动源命令字 [源结构] / the automatic source command
    stHost  : ST_DL_AxisCmd;             // 上位源命令字 [源结构] / the host source command
END_VAR
VAR_OUTPUT
    eWinner     : E_DL_AxisCmdSrc := E_DL_AxisCmdSrc.eNone; // 胜出源 [源] / the winning source
    stWinnerCmd : ST_DL_AxisCmd;                            // 胜出命令字（携带源标签）[源结构] / the winning command carrying its label
    bAnyActive  : BOOL := FALSE;                            // 存在任一源请求 [-] / any source requests
    bSwitched   : BOOL := FALSE;                            // 源切换单拍脉冲 [-] / the source switch one shot pulse
    bError      : BOOL := FALSE;                            // 故障锁存位 [-] / the latched fault bit
    eErr        : UDINT := 16#0000_0000;                    // 错误码，0 = 正常 / the error code, zero is ok
END_VAR
VAR
    _bInit     : BOOL := FALSE;                                // 首拍初始化标志（R310）/ the first scan flag
    _eWinner   : E_DL_AxisCmdSrc := E_DL_AxisCmdSrc.eNone;     // 胜出源副本，段 6 单点映射 / the winning source copy
    _ePrev     : E_DL_AxisCmdSrc := E_DL_AxisCmdSrc.eNone;     // 上拍胜出源（切换沿判据，保持型不入预清，FB32-1）/ the previous winner, held across the scans
    _stWin     : ST_DL_AxisCmd;                                // 胜出命令字副本 / the winning command copy
    _bSwitched : BOOL := FALSE;                                // 切换单拍内部位，段 1 预清段 6 映射 / the internal switch bit, preset then mapped
    _bNoneReq  : BOOL := FALSE;                                // 本拍无源请求标记（逐拍重算）[-] / the no request flag, recomputed every scan
    _bNonFin   : BOOL := FALSE;                                // 胜出命令非有限标记（逐拍重算）[-] / the non finite winner flag, recomputed every scan
    _bFault    : BOOL := FALSE;                                // 故障锁存位（非有限降级置位，复位沿清除，D2 返修）/ the fault latch bit, set on the degrade and cleared by the reset edge
    rtReset    : R_TRIG;                                       // 复位沿实例，段 0 无条件刷新（D2 返修新增）/ the reset edge instance, refreshed unconditionally
END_VAR

// 段 0｜复位沿无条件周期刷新（禁入分支，R7；D2 返修新增）/ segment 0, the unconditional refresh of the reset edge
rtReset(CLK := bReset); // 故障复位沿 / the fault reset edge

// 段 1｜首拍初始化与单拍标志预清（仅单拍标志入清单，R32 FB32-1；R256）/ segment 1, the first scan init and the one shot preset
IF rtReset.Q THEN // 复位沿：清故障锁存（解除路径：复位沿恒可达，R152 自证）/ the reset edge clears the fault latch, the release path is reachable
    _bFault := FALSE; // 清故障锁存 / clear the fault latch
END_IF
IF NOT _bInit THEN // 首拍一拍 / the first scan
    _bInit := TRUE; // 置首拍标志 / raise the first scan flag
    _eWinner := E_DL_AxisCmdSrc.eNone; // 胜出源显式落无源 / place the winner to none explicitly
    _ePrev := E_DL_AxisCmdSrc.eNone; // 上拍源显式落无源 / place the previous winner to none explicitly
END_IF
_bSwitched := FALSE; // 切换脉冲预清零 / preset the switch pulse false
_bNoneReq := FALSE; // 无源标记预清零 / preset the no request flag false
_bNonFin := FALSE; // 非有限标记预清零 / preset the non finite flag false

// 段 2｜优先级仲裁（每拍全量重判，数值小者优先，边界二）/ segment 2, the priority arbitration recomputed every scan
_eWinner := E_DL_AxisCmdSrc.eNone; // 胜出源先置无源 / preset the winner to none
IF bEnable AND (stSafe.eSrc = E_DL_AxisCmdSrc.eSafe) THEN // 安全源请求且标签自洽 / the safety source requests with its own label
    _eWinner := E_DL_AxisCmdSrc.eSafe; // 安全源胜出（最高优先级）/ the safety source wins
ELSIF bEnable AND (stJog.eSrc = E_DL_AxisCmdSrc.eJog) THEN // 手动源请求 / the jog source requests
    _eWinner := E_DL_AxisCmdSrc.eJog; // 手动源胜出 / the jog source wins
ELSIF bEnable AND (stAuto.eSrc = E_DL_AxisCmdSrc.eAuto) THEN // 自动源请求 / the automatic source requests
    _eWinner := E_DL_AxisCmdSrc.eAuto; // 自动源胜出 / the automatic source wins
ELSIF bEnable AND (stHost.eSrc = E_DL_AxisCmdSrc.eHost) THEN // 上位源请求 / the host source requests
    _eWinner := E_DL_AxisCmdSrc.eHost; // 上位源胜出 / the host source wins
END_IF
IF _eWinner = E_DL_AxisCmdSrc.eNone THEN // 无源请求（含失能）/ no source requests or disabled
    _bNoneReq := TRUE; // 置无源标记 / raise the no request flag
END_IF

// 段 3｜胜出命令字整份搬运（携带源标签，边界三；CASE 逐源取，ELSE 兜零命令）/ segment 3, the winning command transfer with the source label
CASE _eWinner OF
    E_DL_AxisCmdSrc.eSafe: // 安全源 / the safety source
        _stWin := stSafe; // 整份搬运 / transfer the whole structure
        _stWin.eSrc := E_DL_AxisCmdSrc.eSafe; // 源标签归一（防调用方填错）/ normalise the label against a caller mistake
    E_DL_AxisCmdSrc.eJog: // 手动源 / the jog source
        _stWin := stJog; // 整份搬运 / transfer the whole structure
        _stWin.eSrc := E_DL_AxisCmdSrc.eJog; // 源标签归一 / normalise the label
    E_DL_AxisCmdSrc.eAuto: // 自动源 / the automatic source
        _stWin := stAuto; // 整份搬运 / transfer the whole structure
        _stWin.eSrc := E_DL_AxisCmdSrc.eAuto; // 源标签归一 / normalise the label
    E_DL_AxisCmdSrc.eHost: // 上位源 / the host source
        _stWin := stHost; // 整份搬运 / transfer the whole structure
        _stWin.eSrc := E_DL_AxisCmdSrc.eHost; // 源标签归一 / normalise the label
    ELSE // 无源或非法枚举值：零命令（安全侧，边界五）/ none or an illegal value, the zero command
        _stWin.eSrc := E_DL_AxisCmdSrc.eNone; // 标签无源 / the label none
        _stWin.fVelMmS := 0.0; // 速度零 / the zero velocity
        _stWin.fPosMm := 0.0; // 位置零 / the zero position
        _stWin.uFlags := 16#0000_0000; // 标志零 / the zero flags
END_CASE

// 段 4｜胜出命令非有限闸（安全侧零命令，不镜像可能被污染的量，R273）/ segment 4, the non finite gate on the winning command
IF (_stWin.fVelMmS <> _stWin.fVelMmS) OR ((_stWin.fVelMmS - _stWin.fVelMmS) <> (_stWin.fVelMmS - _stWin.fVelMmS)) THEN // 速度非有限 / the velocity is not finite
    _bNonFin := TRUE; // 置非有限标记 / raise the non finite flag
END_IF
IF (_stWin.fPosMm <> _stWin.fPosMm) OR ((_stWin.fPosMm - _stWin.fPosMm) <> (_stWin.fPosMm - _stWin.fPosMm)) THEN // 位置非有限 / the position is not finite
    _bNonFin := TRUE; // 置非有限标记 / raise the non finite flag
END_IF
IF _bNonFin THEN // 非有限：降级为零命令 / degrade to the zero command
    _bFault := TRUE; // 锁存故障（D2：故障级码锁存至复位沿，R187）/ latch the fault until the reset edge
    _eWinner := E_DL_AxisCmdSrc.eNone; // 胜出源同步落无源（D1：降级双通道一致，R283）/ sink the winner to none in step with the label
    _stWin.eSrc := E_DL_AxisCmdSrc.eNone; // 标签降级（不再宣称来源）/ degrade the label
    _stWin.fVelMmS := 0.0; // 速度零 / the zero velocity
    _stWin.fPosMm := 0.0; // 位置零 / the zero position
    _stWin.uFlags := 16#0000_0000; // 标志零 / the zero flags
END_IF

// 段 5｜源切换沿判据（保持型上拍源，边界四）/ segment 5, the source switch edge
IF _eWinner <> _ePrev THEN // 与上拍胜出源不同 / differs from the previous winner
    _bSwitched := TRUE; // 置切换单拍 / raise the switch pulse
END_IF
_ePrev := _eWinner; // 上拍源快照（主体末行赋值，跨拍保持）/ snapshot the winner at the body end

// 段 6｜统一出口（内部副本单点映射，R180；故障码回放，R187）/ segment 6, the unified outlet
eWinner := _eWinner; // 胜出源出口 / the winner outlet
stWinnerCmd := _stWin; // 胜出命令字出口 / the winning command outlet
bAnyActive := NOT _bNoneReq; // 有源请求出口 / the any request outlet
bSwitched := _bSwitched; // 切换单拍出口 / the switch pulse outlet
IF _bFault THEN // 故障锁存回放优先（D2：锁存至复位沿，R187）/ the latched fault replays first until the reset edge
    bError := TRUE; // 故障锁存位出口（与 _bFault 同源，R191）/ the fault outlet from the same latch
    eErr := 16#0004_0622; // 故障级：胜出命令含非有限量（锁存回放）/ fault grade, a non finite command quantity, replayed
ELSIF _bNoneReq THEN // 无源请求 / no request
    bError := FALSE; // 无故障 / no fault
    eErr := 16#0004_0620; // 信息级：无任何命令源请求 / informational, no source requests
ELSIF _bSwitched THEN // 源切换 / a source switch
    bError := FALSE; // 无故障 / no fault
    eErr := 16#0004_0621; // 信息级：发生源切换 / informational, a source switch happened
ELSE // 无事件 / no event
    bError := FALSE; // 无故障 / no fault
    eErr := 16#0000_0000; // 正常 / ok
END_IF
END_FUNCTION_BLOCK
